(* IEC 61131-3 sources: plcassist-cli/packages/volt-lsp-iec/test-corpus/pro2193/Device/Plc Logic/Application/09 Misc/Library Manager/L_TT1P_TechnologyModules (part 3) *)

(* ---- L_MB1P_MOVEPICKANDPLACEBASE.fb ---- *)
FUNCTION_BLOCK L_MB1P_MOVEPICKANDPLACEBASE EXTENDS L_MC4P_Template_AG_KIN
VAR_INPUT
	DWCYCLESTAMP : DWORD;
	XEXECUTE : BOOL;
	XABORT : BOOL;
	WMOVEMODE : WORD;
	XFULLPATHBLENDING : BOOL;
	XNOTCOORDINATEDSTOPALL : BOOL;
	ETARGETCOORDSYSTEM : L_MC4P_CoordSystem;
	ESTARTCOORDSYSTEM : L_MC4P_CoordSystem;
	LRSTARTBLENDINGRADIUS : LREAL;
	EBUFFERMODE : MC_BUFFER_MODE := MC_BUFFER_MODE.mcBlendingLow;
	LRPATHJERK : LREAL := 1E+24;
	LRGRIPPERTIME : LREAL;
	XPULSEGRIPPERINTERRUPT : BOOL;
	XCALCPROFILEMOVEPATH : BOOL;
	WCONVEYOREXTRAPOLMODE : WORD;
	LRCONVEYOREXTRAPOLOFFSET : LREAL;
	LRCONVEYOREXTRAPOLVEL : LREAL;
	LRCONVEYOREXTRAPOLTIME : LREAL;
	XGETOVERRIDEFADINGTIME : BOOL;
END_VAR
VAR_OUTPUT
	XERROR : BOOL;
	XWARNING : BOOL;
	EERRORID : L_IE1P_Error;
	XBUSY : BOOL;
	XDONE : BOOL;
	XPROFILEINPREPARATION : BOOL;
	XCOMMANDABORTED : BOOL;
	XACTIVE : BOOL;
	XPATHHOLD : BOOL;
	XPATHHOLDONGRIPPERPOINT : BOOL;
	ESETSEGMENTTYPEOUT : L_MC4P_SegmentType;
	ALRTARGETPOSWCSOUT : ARRAY [1..6] OF LREAL;
	ALRTARGETPOSAUXOUT : ARRAY [1..6] OF LREAL;
	XPULSEGRIPPER : BOOL;
	WPATHMODEOUT : WORD;
	ITARGETPOINT : SINT;
	INUMOFSEGMENTSINPROFILE : SINT;
	XSETPATHPREPARATIONTIMEVALID : BOOL;
	LRSETPATHPREPARATIONTIMEOUT : LREAL;
	LRSETPROFILEIPOTIMEOUT : LREAL;
	XPRECALCPROFILERESTTIMEVALID : BOOL;
	LRPRECALCPROFILERESTTIME : LREAL;
	LRPRECALCPROFILEORIRESTTIME : LREAL;
	XUPDATEPROFILESYNCRESTTIME : BOOL;
	XPRECALCPROFILESYNCRESTTIME : BOOL;
	LRPRECALCPROFILESYNCRESTTIME : LREAL;
	XPRECALCPROFILESYNCOUTTIME : BOOL;
	LRPRECALCPROFILESYNCOUTTIME : LREAL;
	LRPRECALCPROFILETIME : LREAL;
	LRINTERRUPTPATHACC : LREAL;
	XIPOTIMEMOVEFROMTARGETVALID : BOOL;
	WIPOTIMEMOVEFROMTARGETCVNO : WORD;
	LRIPOTIMEMOVEFROMTARGET : LREAL;
	LRCONVEYOREXTRAPOLOFFSETOUT : LREAL;
	XPARVALID : BOOL := FALSE;
	LROVERRIDEFADINGTIME : LREAL;
	LRMAXVEL : LREAL := 10;
	LRMAXACC : LREAL := 100;
	LRMAXDEC : LREAL := 100;
	LRMAXJERK : LREAL := 100;
	XRESERVEFUNID : BOOL;
	XWAITDISABLEMOVECONTPATH : BOOL;
END_VAR
VAR_IN_OUT
	MC_MOVELINABSCONTINUEPROFILE : L_MC4P_MoveLinearAbsolute_Internal;
END_VAR
VAR
	WMOVEMODE_INT : WORD;
	XSINGLESTEP_INT : BOOL;
	XPULSEGRIPPERINTERRUPT_INT : BOOL;
	LRSTARTBLENDINGRADIUS_INT : LREAL;
	ICONTPGRIPPERINTERRUPT_INT : INT;
	XINTERRUPTONGRIPPERPOINTATMODE_INT : BOOL;
	LRPRECALCPROFILERESTTIME_INT : LREAL;
	LRSETPROFILEIPOTIME_INT : LREAL;
	LRACTTIMEOR : LREAL;
	LRSYNCRONISEDTIME : LREAL;
	LRACTSYNCRONISEDTIME : LREAL;
	XACTSYNCRONISEDTIMEOLDVALID : BOOL;
	LRACTSYNCRONISEDTIME_OLD : LREAL;
	XRESETSUPERPOSONCV_INT : BOOL;
	LRSYNCINZDISTFACTOR_INT : LREAL := 0.5;
	LRSYNCINDISTFACTOR_INT : LREAL := 1;
	LRSYNCOUTDISTFACTOR_INT : LREAL := 1;
	LRWAITTIMESTATICTARGETPOS_INT : LREAL;
	XINTERRUPTATSTATICTARGETPOS_INT : BOOL;
	XINTERRUPTATTARGETONCV_INT : BOOL;
	XABORTACTIVE : BOOL;
	WMODE_OLD : WORD;
	WMODE_INT : WORD;
	LRADDPROFILERESTTIME_INT : LREAL;
	XADDPROFILERESTTIMEVALID : BOOL;
	XACKNTARGETWORKPIECE_INT : BOOL;
	LRAUX1STARTPOS_INT : LREAL;
	XAUX1STARTPOSVALID_INT : BOOL;
	LRASTARTPOS_INT : LREAL;
	XASTARTPOSVALID_INT : BOOL;
	LRBSTARTPOS_INT : LREAL;
	XBSTARTPOSVALID_INT : BOOL;
	LRCSTARTPOS_INT : LREAL;
	XCSTARTPOSVALID_INT : BOOL;
	ETRACKPICKANDPLACETARGET_INT_OLD : L_TT1P_TrackPickAndPlaceTarget;
	ETRACKPICKANDPLACETARGET_INT : L_TT1P_TrackPickAndPlaceTarget;
	EBUFFERMODEINTERNAL_INT : MC_BUFFER_MODE := MC_BUFFER_MODE.mcBlendingLow;
	LWTCHECKSUM_INT : LWORD;
	LRTMPSTARTCOORDSYS : LREAL;
	LRPROFILERESTTIME : LREAL;
	XPRECALCGRIPPERRESTTIMEVALID : BOOL;
	LRPRECALCGRIPPERRESTTIME : LREAL;
	ETRACKPPMOVESTATUS_INT : L_TT1P_TrackPickAndPlaceTargetStatus;
	XPATHHOLD_INT : BOOL;
	XPAHTHOLDDONE_INT : BOOL;
	XPAHTHOLDDONE_LOCK : BOOL;
	REQUESTSINFO : DWORD;
	REQUESTSINFO_OLD : DWORD;
	DWRTRIG : DWORD;
	DWFTRIG : DWORD;
	LRTEMP : LREAL;
	LRTEMP2 : LREAL;
	IDX1 : SINT;
	IDX2 : SINT;
	UIDX : USINT;
	WDX : WORD;
	LRTIME_TMP : LREAL;
	LRALLPOFILETIME : LREAL;
	LRRESTTIMEENDSEGMENT_INT : LREAL;
	IDX_START : SINT;
	IDX_END : SINT;
	XINTERRUPTEDATNEXTBUFFEREDPOS_TMP : BOOL;
	WSTATE : WORD;
	WSTATE_OLD : WORD;
	XSTATEENTRY : BOOL;
	XIPOTIMEMOVEFROMTARGETVALID_OLD : BOOL;
	LRTASKCYCLE : LREAL;
	LRTASKCYCLEOR : LREAL;
	LRTASKCYCLE_INV : LREAL;
	XSTARTPATHLISTISEMPTY : BOOL;
	XCALCPATHPREPARATIONTIME : BOOL;
	XRETURNINIT : BOOL;
	LRTIMECORRFACTORATOR_INT : LREAL;
	LRPRECALCGRIPPERRESTTIMECORROR : LREAL;
	XPRECALCPROFILESYNCOUTTIME_INT : BOOL;
	INUMOFMOVEREL : SINT;
	INUMOFMOVEABS : SINT;
	INUMOFMOVEELLIPTICAL : SINT;
	XEXECUTEAFTERHALT : BOOL;
	INUMOFSEGMENTSEXECUTED : SINT;
	INUMOFMOVERELEXECUTED : SINT;
	INUMOFMOVEABSEXECUTED : SINT;
	INUMOFMOVEELLIPTICALEXECUTED : SINT;
	INUMOFMOVESPLINEEXECUTED : SINT;
	ITARGETPOINTMOVEABS : SINT;
	XNOMOVEFBEXECUTED : BOOL;
	INUMOFMOVEFBSCHECKEDORFEEDINGTIME : SINT;
	LRZSYNCDIST : LREAL;
	EPATHMODE_INT : L_TT1P_PickAndPlacePathMode;
	XGRIPPERCTRLACTIVE_INT : BOOL;
	ISETMOVEFBNOACTIVE : SINT;
	ISETNUMOFMOVEFBSADDTIME : SINT;
	IACKNNUMOFSEGMENTSINPROFILE : SINT;
	IACKNNUMOFMOVEREL : SINT;
	IACKNNUMOFMOVEABS : SINT;
	IACKNNUMOFMOVEELLIPTICAL : SINT;
	INUMOFENABLEDSEGMENTS : SINT;
	XPROFILEINPREPARATION_INT : BOOL;
	XMOVEPROFILEBUSY : BOOL;
	XMOVEPROFILEACTIVE : BOOL;
	XMOVEPROFILEACTIVE_OLD : BOOL;
	XMOVEPROFILEDONE : BOOL;
	XMOVEPROFILENOPULSEGRIPPERDONE : BOOL;
	XMOVEPROFILECOMMANDABORTED : BOOL;
	XMOVEPROFILECOMMANDABORTED_OLD : BOOL;
	XMOVEPROFILEENABLED : BOOL;
	XMOVEPROFILEHOLD : BOOL;
	XHOLDONHALT : BOOL;
	XHOLDONGRIPPERPOINT : BOOL;
	XHOLDONGRIPPERPOINT_OLD : BOOL;
	XMOVEPROFILEERROR : BOOL;
	EMOVEPROFILEERRORID : L_IE1P_Error;
	XMOVEPROFILESTATEINITIAL : BOOL := TRUE;
	ITARGETPOINTOFFSET : INT;
	INUMOFVALIDPROFILETIME : USINT;
	AXPROFILETIMEVALID : ARRAY [1..11] OF BOOL;
	ALRPROFILETIME : ARRAY [1..11] OF LREAL;
	WTARGETMODE_INT : WORD;
	XPRECALCPROFILERESTTIMEVALID_INT : BOOL;
	XPRECALCPROFILERESTTIMEVALID_OLD : BOOL;
	XCONTINUE1STMOVEABSACTIVE : BOOL;
	XCONTINUEPROFILEVIA1STMOVEABS : BOOL;
	XERROR_INVALIDCOORDSYSTEM : BOOL;
	XERRORINVALIDPROFILE : BOOL;
	XERROR_INTERNAL : BOOL;
	IINVALIDEMOVESTATECOUNTER : INT := 0;
	XSETZPOSVALID : BOOL;
	LRSETZPOSITION : LREAL;
	LRSETZPOSITION_OLD : LREAL;
	LRSETZDIST_INT : LREAL;
	LRPATHDIST_INT : LREAL;
	EBUFFERMODEINTERNAL : MC_BUFFER_MODE;
	ETRACKPICKANDPLACETARGET : L_TT1P_TrackPickAndPlaceTarget;
	ETRACKPICKANDPLACETARGET_OLD : L_TT1P_TrackPickAndPlaceTarget;
	ETRACKPPMOVESTATUS : L_TT1P_TrackPickAndPlaceTargetStatus;
	INUMOFACTIVEPATHSEGMENT : INT;
	LRADDPROFILERESTTIME : LREAL;
	LRAUX1STARTPOS : LREAL;
	LRPRECALCINGRIPPERPOSRESTTIME : LREAL;
	LRSYNCINDISTFACTOR : LREAL;
	LRSYNCINZDISTFACTOR : LREAL;
	LRSYNCOUTDISTFACTOR : LREAL;
	LRWAITTIMESTATICTARGETPOS : LREAL;
	LWTCHECKSUM : LWORD;
	WMODE : WORD;
	WMODEOLD : WORD;
	WSTATELINE : WORD;
	XACKNTARGETWORKPIECE : BOOL;
	XGRIPPERCTRLACTIVE : BOOL;
	XGRIPPERSEGMENTTIMEIPOACTIVE : BOOL;
	XINGRIPPERPOS : BOOL;
	XINTERRUPTATSTATICTARGET : BOOL;
	XINTERRUPTATTARGETONCV : BOOL;
	XLASTSEGMENTTIMEIPOACTIVE : BOOL;
	XPATHHOLDONENDHALT : BOOL;
	XPRECALCINGRIPPERPOSRESTTIMEVALID : BOOL;
	XRESETSUPERPOSONCV : BOOL;
	XRTRIGIPOTIMEMOVEFROMTARGETVALID : BOOL;
END_VAR
END_FUNCTION_BLOCK

METHOD ABORT
END_METHOD

METHOD CALL_ABORTINPUT
END_METHOD

METHOD CALL_ALLOCPOINTADR
END_METHOD

METHOD CALL_CALCTIME
END_METHOD

METHOD CALL_CHECKSTATEENTRY
END_METHOD

METHOD CALL_DISABLEMOVECONTPATH
VAR_IN_OUT
	AXESGROUP : AXES_GROUP_KIN;
END_VAR
END_METHOD

METHOD CALL_ERRORHANDLER
END_METHOD

METHOD CALL_FBMETHODS
END_METHOD

METHOD CALL_FBMETHODS_MOVEFBS
END_METHOD

METHOD CALL_GRIPPERCONTROL
END_METHOD

METHOD CALL_MC_MOVELINABS
VAR_IN_OUT
	AXESGROUP : AXES_GROUP_KIN;
END_VAR
END_METHOD

METHOD CALL_MC_MOVELINABS_1STCONTINUEPROFILE
VAR_IN_OUT
	AXESGROUP : AXES_GROUP_KIN;
END_VAR
END_METHOD

METHOD CALL_OUTPUT
END_METHOD

METHOD CALL_OUTPUTDISABLED
END_METHOD

METHOD CALL_PROFILE_STATUS
END_METHOD

METHOD CALL_PROFILE_STATUS_1STCONTINUEPROFILE
END_METHOD

METHOD CALL_PROFILE_STATUS_INIT
END_METHOD

METHOD CALL_PROFILE_STATUS_OUTPUT
END_METHOD

METHOD CALL_REQUESTS_EXT
END_METHOD

METHOD CALL_RESET
END_METHOD

METHOD CALL_RESETCOMMANDS
END_METHOD

METHOD CALL_RESETOUTPUT
END_METHOD

METHOD CALL_RESETTEMPMEMORY
END_METHOD

METHOD CALL_STATEMACHINE
END_METHOD

METHOD GET_LRPRECALCPROFILERESTTIMEFASTSYNCOUT : LREAL
END_METHOD

METHOD GET_LRRESTTIMEBEVOREMOVETOPARKPOS : LREAL
END_METHOD

METHOD GET_LRPROFILETIMEZTARGETDIST : BOOL
VAR_IN_OUT
	XPROFILETIMEZTARGETDISTVALID : BOOL;
	LRPROFILETIMEZTARGETDIST : LREAL;
END_VAR
END_METHOD

METHOD SET_EXTERNALGRIPPERTRIGGER
END_METHOD

METHOD CALL_EMPTY
END_METHOD

METHOD CALL_CONTINUEPROFILE
END_METHOD

METHOD CALL_CONTINUEPROFILE1STBLENDING
END_METHOD

METHOD CALL_CONTINUEPROFILE_MOVEABSCONTINUEPROFILE
END_METHOD

METHOD CALL_DATAFROMIPOLISTELEMENT
END_METHOD

METHOD CALL_DATAFROMIPOLISTELEMENTATSTOP
END_METHOD

METHOD CALL_DISABLEMOVEFBS
END_METHOD

METHOD CALL_EXECUTEPROFILE
END_METHOD

METHOD CALL_LOCKPAR
END_METHOD

METHOD CALL_READSTARTPOSITION
END_METHOD

METHOD CALL_SETPROFILE
END_METHOD

METHOD FUN_GETOVERRIDEFADINGTIME
VAR_INPUT
	INUMOFMOVEFBS : SINT;
END_VAR
END_METHOD

METHOD GET_PROFILETIME_MOVELINABSCONTINUEPROFILE : LREAL
END_METHOD

METHOD RESET_PRECALCPROFILETIME
END_METHOD

METHOD SET_TONEXTSEGMENTAFTERPATHHOLD
END_METHOD

METHOD CALL_INIT
END_METHOD

METHOD CALL_S000_CYCLIC
END_METHOD

(* ---- L_MB1P_MOVEPICKANDPLACEBASEEXTENDED.fb ---- *)
FUNCTION_BLOCK L_MB1P_MOVEPICKANDPLACEBASEEXTENDED EXTENDS L_MB1P_MovePickAndPlaceBase
VAR_INPUT
	ALRTARGETPOS : ARRAY [1..12] OF LREAL;
	LRZSTARTDIST : LREAL;
	LRZTARGETDIST : LREAL;
	LRVELFACTORATTARGET : LREAL := 1;
	LRACCDECFACTORATTARGET : LREAL := 1;
	XZSTARTDISTTOPARKPOS : BOOL;
	LRZSTARTDISTTOPARKPOS : LREAL;
	XZTARGETDISTFROMPARKPOS : BOOL;
	LRZTARGETDISTFROMPARKPOS : LREAL;
	LRBLENDINGRADIUS : LREAL;
	LRPATHVEL : LREAL := 10;
	LRPATHACC : LREAL := 100;
	LRPATHDEC : LREAL := 100;
	EORIENTATIONMODE : L_MC4P_Orientation_Mode := L_MC4P_Orientation_Mode.ShortestSpacialWay;
	EADIRECTION : MC_DIRECTION := MC_DIRECTION.mcShortestWay;
	EBDIRECTION : MC_DIRECTION := MC_DIRECTION.mcShortestWay;
	ECDIRECTION : MC_DIRECTION := MC_DIRECTION.mcShortestWay;
END_VAR
VAR_IN_OUT
	MC_MOVELINREL : L_MC4P_MoveLinearRelative_Internal;
	AMC_MOVELINABS : ARRAY [1..2] OF L_MC4P_MoveLinearAbsolute_Internal;
END_VAR
VAR
	LRZSTARTDIST_INT : LREAL;
	LRZTARGETDIST_INT : LREAL;
	LRZDISTELLIPTICAL_INT : LREAL;
	LRZSTARTPOSWCS_INT : LREAL;
	LRZTARGETPOSWCS_INT : LREAL;
	LRZSTARTPOSINTARGET : LREAL;
	LRZTARGETPOSINTARGET : LREAL;
	LRPRECALCPROFILETIMEINTARGETCOORDSYSTEM : LREAL;
	LRPRECALCPROFILETIMEZTARGETDIST : LREAL;
	XCALCPRECALCPROFILETIMEZTARGETDIST : BOOL := FALSE;
	WPROFILEMASK_LOCK : WORD;
	WPROFILEMODE_LOCK : WORD;
	LRZDIST_INT : LREAL;
	XLASTSEGMENTTIMEIPOACTIVE : BOOL;
END_VAR
END_FUNCTION_BLOCK

METHOD CALL_CALCTIME
END_METHOD

METHOD CALL_DISABLEMOVECONTPATH
VAR_IN_OUT
	AXESGROUP : AXES_GROUP_KIN;
END_VAR
END_METHOD

METHOD CALL_FBMETHODS_MOVEFBS
END_METHOD

METHOD CALL_MC_MOVELINABS
VAR_IN_OUT
	AXESGROUP : AXES_GROUP_KIN;
END_VAR
END_METHOD

METHOD CALL_MC_MOVELINREL
VAR_IN_OUT
	AXESGROUP : AXES_GROUP_KIN;
END_VAR
END_METHOD

METHOD CALL_OUTPUTDISABLED
END_METHOD

METHOD CALL_PROFILE_STATUS
END_METHOD

METHOD CALL_PROFILE_STATUS_MOVEABS
END_METHOD

METHOD CALL_PROFILE_STATUS_MOVEREL
END_METHOD

METHOD CALL_PROFILE_STATUS_OUTPUT
END_METHOD

METHOD CALL_RESETCOMMANDS
END_METHOD

METHOD CALL_CONTINUEPROFILE
END_METHOD

METHOD CALL_CONTINUEPROFILE_MOVEABS
END_METHOD

METHOD CALL_CONTINUEPROFILE_MOVEREL
END_METHOD

METHOD CALL_DATAFROMIPOLISTELEMENTATSTOP
END_METHOD

METHOD CALL_DISABLEMOVEFBS
END_METHOD

METHOD CALL_EXECUTEPROFILE
END_METHOD

METHOD CALL_LOCKPAR
END_METHOD

METHOD CALL_LOCKPAR_ZDIST
END_METHOD

METHOD CALL_LOCKPAR_ZSTARTDISTTOPARKPOS
END_METHOD

METHOD CALL_LOCKPAR_ZTARGETDISTFROMPARKPOS
END_METHOD

METHOD CALL_SETPROFILE
END_METHOD

METHOD CALL_SETPROFILE_TOFIRSTPOINT
END_METHOD

METHOD GET_PROFILETIME_MOVELINREL : LREAL
END_METHOD

METHOD GET_PROFILETIME_AMOVEABS : LREAL
VAR_IN_OUT
	IFBNO : SINT;
END_VAR
END_METHOD

METHOD SET_TONEXTSEGMENTAFTERPATHHOLD
END_METHOD

(* ---- L_MB1P_MOVEPICKANDPLACEELLIPTICAL.fb ---- *)
FUNCTION_BLOCK L_MB1P_MOVEPICKANDPLACEELLIPTICAL EXTENDS L_MB1P_MovePickAndPlaceBaseExtended
VAR_INPUT
	EPATHMODE : L_TT1P_PickAndPlacePathMode;
	LRZDISTELLIPTICAL : LREAL;
	XZSTARTPOSMCS : LREAL;
	LRZSTARTPOSWCS : LREAL;
	LRZTARGETPOSWCS : LREAL;
	ALRDIRECTIONTOPARKPOS : ARRAY [1..3] OF LREAL := [0, 0, 1];
	ALRDIRECTIONFROMPARKPOS : ARRAY [1..3] OF LREAL := [0, 0, 1];
END_VAR
VAR_IN_OUT
	FB_MOVEELLIPTICAL : L_MC4P_MoveEllipticalAbsolutePnP_Internal;
END_VAR
VAR
	XTEST : BOOL;
	XUSEORICAM_INT : BOOL;
	LRAUX1CAMTARGETPOS : LREAL;
	LRCCAMTARGETPOS : LREAL;
	XLASTSEGMENTTIMEIPOACTIVE : BOOL;
	XUSEORICAM : BOOL;
END_VAR
END_FUNCTION_BLOCK

METHOD CALL_DISABLEMOVECONTPATH
VAR_IN_OUT
	AXESGROUP : AXES_GROUP_KIN;
END_VAR
END_METHOD

METHOD CALL_FBMETHODS_MOVEFBS
END_METHOD

METHOD CALL_FB_MOVEELLIPTICAL
VAR_IN_OUT
	AXESGROUP : AXES_GROUP_KIN;
END_VAR
END_METHOD

METHOD CALL_OUTPUTDISABLED
END_METHOD

METHOD CALL_PROFILE_STATUS
END_METHOD

METHOD CALL_PROFILE_STATUS_MOVEELLIPTICAL
END_METHOD

METHOD CALL_RESETCOMMANDS
END_METHOD

METHOD GET_LRPROFILETIMEZTARGETDIST : BOOL
VAR_IN_OUT
	XPROFILETIMEZTARGETDISTVALID : BOOL;
	LRPROFILETIMEZTARGETDIST : LREAL;
END_VAR
END_METHOD

METHOD CALL_CONTINUEPROFILE
END_METHOD

METHOD CALL_CONTINUEPROFILE_MOVEELLIPTICAL
END_METHOD

METHOD CALL_DATAFROMIPOLISTELEMENTATSTOP
END_METHOD

METHOD CALL_DISABLEMOVEFBS
END_METHOD

METHOD CALL_EXECUTEPROFILE
END_METHOD

METHOD CALL_LOCKPAR
END_METHOD

METHOD CALL_LOCKPAR_ZDIST
END_METHOD

METHOD CALL_LOCKPAR_ZSTARTDISTTOPARKPOS
END_METHOD

METHOD CALL_LOCKPAR_ZTARGETDISTFROMPARKPOS
END_METHOD

METHOD CALL_SETPROFILE
END_METHOD

METHOD CALL_SETPROFILE_TOFIRSTPOINTEXTENDEDELLIPTICAL
END_METHOD

METHOD GET_PATHLENGTH_MOVEELLIPTICAL : LREAL
END_METHOD

METHOD GET_PROFILETIME_MOVEELLIPTICAL : LREAL
END_METHOD

(* ---- L_MB1P_MOVEPICKANDPLACESTATE.fb ---- *)
FUNCTION_BLOCK L_MB1P_MOVEPICKANDPLACESTATE EXTENDS L_MB1P_MovePickAndPlaceBase
VAR_INPUT
	XINTERRUPTONGRIPPERPOINT : BOOL;
	XSHIFTEXECUTENEXTPROFILE : BOOL;
	LRPATHPREPARATIONTIME : LREAL;
	XSTARTPOINTINHALT : BOOL;
	XHOLDMOVEPATH : BOOL;
	IPOINTNOSYNCIN : SINT;
	IPOINTNOPULSEGRIPPER : SINT;
	XACKPATHHALT : BOOL;
	XEXECUTEPROFILEAFTERGRIPPER : BOOL;
END_VAR
VAR_OUTPUT
	XPATHINTERRUPTOUT : BOOL;
	ETARGETCOORDSYSTEMOUT : L_MC4P_CoordSystem;
	ALRTARGETPOS : ARRAY [1..12] OF LREAL;
	ALRINTERMEDIANTEPOINT : ARRAY [1..12] OF LREAL;
	LRENDBLENDINGRADIUS : LREAL;
	XENDHALT : BOOL;
	XEXECUTEDPROFILEAFTERGRIPPER : BOOL;
END_VAR
VAR_IN_OUT
	ASCPROFILEPAR : ARRAY [1..10] OF L_TT1P_scProfilePar;
	AMC_MOVELINABS : ARRAY [1..10] OF L_MC4P_MoveLinearAbsolute_Internal;
END_VAR
VAR
	LRPATHPREPARATIONTIME_INT : LREAL;
	XSHIFTEXECUTENEXTPROFILE_INT : BOOL;
	XWAITOFNEXTPROFILE_INT : BOOL;
	WWAITOFNEXTPROFILECNTR : WORD;
	XNEXTPROFILEWAITFOREXECUTE_INT : BOOL;
	XEXECUTEPROFILEAFTERGRIPPER_LOCK : BOOL;
	XINTERRUPTONGRIPPERPOINT_INT : BOOL;
	XINTERRUPTONGRIPPERPOINT_OLD : BOOL;
	XINGRIPPERPOS_INT : BOOL;
	XINSYNCPOS_INT : BOOL;
	LRENDPATHVEL_INT : LREAL;
	LRENDPATHACC_INT : LREAL;
	LRENDPATHDEC_INT : LREAL;
	INUMOFMOVEABSEXECUTEDAFTERHALT : SINT;
	IRETURNINITCNTR : INT;
	XREADSTARTPOSACTIVE : BOOL;
	XIPOTIMEMOVEFROMTARGETACTIVE_INT : BOOL;
	ICNTRACKPATHHALT_INT : INT;
	ICNTRACKPATHHALTREST_INT : INT;
	ICNTRACKPATHHALTFORGRIPPER_INT : INT;
	ICNTRACKPATHHALT_LOCK : INT;
	INUMOFHALTINPROFILE_INT : INT;
	IPOINTNOSYNCOUT_INT : SINT;
	IPOINTNOSYNCIN_INT : SINT;
	IPOINTNOPULSEGRIPPER_INT : SINT;
	ALRSTARTPOS_INT : ARRAY [1..6] OF LREAL;
	ECOORDSYSTEMP1START : L_MC4P_CoordSystem;
	ECOORDSYSTEMP2ACT : L_MC4P_CoordSystem;
	ECOORDSYSTEMP3NEXT : L_MC4P_CoordSystem;
	ALRP1START : ARRAY [1..3] OF LREAL;
	ALRP2ACT : ARRAY [1..3] OF LREAL;
	ALRP3NEXT : ARRAY [1..3] OF LREAL;
	XPOINTSONASTRAIGHTLINE : BOOL;
	XNOFUNKTION : BOOL;
	XSTARTPOSVALID_INT : BOOL;
	XPROFILEEXECUTED_INT : BOOL;
	XEXECUTENEXTMOVEPP_INT : BOOL;
	XACKENDHALT_INT : BOOL;
	AXHALT : ARRAY [0..10] OF BOOL;
	AITARGETPOINTOFFSETATMOVEABS : ARRAY [0..10] OF INT;
	AXMOVELINABSACTIVE : ARRAY [0..10] OF BOOL;
	XVALIDSYNCRESTTIME_OLD : BOOL;
	XVALIDSYNCRESTTIME_INT : BOOL;
	XVALIDSYNCOUTRESTTIME_OLD : BOOL;
	XVALIDSYNCOUTRESTTIME_INT : BOOL;
	LRRESTTIMESYNC_INT : LREAL;
	LRRESTTIMESYNCOUT_INT : LREAL;
	XVALIDPULSEGRIPPERRESTTIME_OLD : BOOL;
	XVALIDPULSEGRIPPERRESTTIME_INT : BOOL;
	LRPULSEGRIPPERRESTTIME_INT : LREAL;
	LRBLENDINGRADIUS_TMP : LREAL;
	XCALCDIST_TMP : BOOL;
	XCALCINTERMEDIANTEPOINT : BOOL;
	AXCALCPATHLEGTHBETWEENPOINTS : ARRAY [0..10] OF BOOL;
	ALRPATHLENGTHBETWEENPOINTS : ARRAY [0..10] OF LREAL;
	ALRAUX1POINTS : ARRAY [0..10] OF LREAL;
	ALRAPOINTS : ARRAY [0..10] OF LREAL;
	ALRBPOINTS : ARRAY [0..10] OF LREAL;
	ALRCPOINTS : ARRAY [0..10] OF LREAL;
	IFORCNT : SINT;
	XCALC999AUX1TARGETPOS : BOOL;
	XCALC999ATARGETPOS : BOOL;
	XCALC999BTARGETPOS : BOOL;
	XCALC999CTARGETPOS : BOOL;
	IFIRSTPOINTATPROFILEPAR : SINT;
	ILISTELEMENTATSTOPCNTR_INT : SINT;
	XNEXTPROFILEPOINTATBLENDING_INT : BOOL;
	MC_GROUPREADACTUALPOSITION1 : MC_GroupReadActualPosition;
	ALRPROFILESTARTPOS : ARRAY [1..6] OF LREAL;
	ILISTELEMENTATSTOPCNTR : SINT;
	LRENDPATHACC : LREAL;
	LRENDPATHDEC : LREAL;
	LRENDPATHVEL : LREAL;
	WSTATELINE : WORD;
	XEXECUTENEXTMOVEPP : BOOL;
	XGRIPPERSEGMENTTIMEIPOACTIVE : BOOL;
	XINGRIPPERPOS : BOOL;
	XLASTSEGMENTTIMEIPOACTIVE : BOOL;
	XMOVEFROMTARGETACTIVE : BOOL;
	XNEXTPROFILEPOINTATBLENDING : BOOL;
	XNEXTPROFILEWAITFOREXECUTE : BOOL;
	XPATHHOLDONENDHALT : BOOL;
END_VAR
END_FUNCTION_BLOCK

METHOD CALL_ABORTINPUT
END_METHOD

METHOD CALL_CALCTIME
END_METHOD

METHOD CALL_DISABLEMOVECONTPATH
VAR_IN_OUT
	AXESGROUP : AXES_GROUP_KIN;
END_VAR
END_METHOD

METHOD CALL_ERRORHANDLER
END_METHOD

METHOD CALL_FBMETHODS
END_METHOD

METHOD CALL_FBMETHODS_MOVEFBS
END_METHOD

METHOD CALL_MC_GROUPREADACTUALPOSITION
END_METHOD

METHOD CALL_MC_MOVELINABS
VAR_IN_OUT
	AXESGROUP : AXES_GROUP_KIN;
END_VAR
END_METHOD

METHOD CALL_OUTPUT
END_METHOD

METHOD CALL_OUTPUTDISABLED
END_METHOD

METHOD CALL_PROFILE_STATUS
END_METHOD

METHOD CALL_PROFILE_STATUS_MOVEABS
END_METHOD

METHOD CALL_PROFILE_STATUS_INIT
END_METHOD

METHOD CALL_PROFILE_STATUS_OUTPUT
END_METHOD

METHOD CALL_REQUESTS_EXT
END_METHOD

METHOD CALL_RESETCOMMANDS
END_METHOD

METHOD CALL_RESETOUTPUT
END_METHOD

METHOD GET_LRPRECALCPROFILERESTTIMEFASTSYNCOUT : LREAL
END_METHOD

METHOD GET_LRRESTTIMEBEVOREMOVETOPARKPOS : LREAL
END_METHOD

METHOD GET_IACKPATHHALTCNTRREST
VAR_IN_OUT
	ICOUNTER : INT;
END_VAR
END_METHOD

METHOD CALL_CALC999TARGETPOS
VAR_INPUT
	IPOINTNO : SINT;
END_VAR
VAR_IN_OUT
	ALRPOINTS : ARRAY [0..10] OF LREAL;
	ALRLEGTHBETWEENPOINTS : ARRAY [0..10] OF LREAL;
END_VAR
END_METHOD

METHOD CALL_CHECKORIDIRECTION_SWITCHTOSHORTESTWAY
VAR_INPUT
	LRCYCLELENGTH : LREAL;
	LRPOSSTART : LREAL;
	LRPOSEND : LREAL;
	EDIRECTION : MC_DIRECTION;
END_VAR
VAR_OUTPUT
	EDIRECTIONOUT : MC_DIRECTION;
END_VAR
END_METHOD

METHOD CALL_CONTINUEPROFILE
END_METHOD

METHOD CALL_CONTINUEPROFILE_MOVEABS
END_METHOD

METHOD CALL_DATAFROMIPOLISTELEMENTATSTOP
END_METHOD

METHOD CALL_DISABLEMOVEFBS
END_METHOD

METHOD CALL_EXECUTEPROFILE
END_METHOD

METHOD CALL_LOCKPAR
END_METHOD

METHOD CALL_READSTARTPOSITION
END_METHOD

METHOD CALL_SETPROFILE
END_METHOD

METHOD FUN_POINTSONASTRAIGHTLINE : BOOL
VAR_OUTPUT
	XNOFUNKTION : BOOL;
END_VAR
VAR_IN_OUT
	AXESGROUP : AXES_GROUP_KIN;
	ALRP1 : ARRAY [1..3] OF LREAL;
	ECOORDSYSTEMP1 : L_MC4P_CoordSystem;
	ALRP2 : ARRAY [1..3] OF LREAL;
	ECOORDSYSTEMP2 : L_MC4P_CoordSystem;
	ALRP3 : ARRAY [1..3] OF LREAL;
	ECOORDSYSTEMP3 : L_MC4P_CoordSystem;
END_VAR
END_METHOD

METHOD GET_FIRSTPROFILEPOINTPAR
VAR_IN_OUT
	SCPROFILEPAR : L_TT1P_scProfilePar;
END_VAR
END_METHOD

METHOD GET_INUMOFACTIVEHALTPOINTS : INT
END_METHOD

METHOD GET_PROFILETIME_AMOVEABS : LREAL
VAR_IN_OUT
	IFBNO : SINT;
END_VAR
END_METHOD

METHOD SET_ACKENDHALT
END_METHOD

METHOD SET_FIRSTPROFILEPOINTATBLENDING
VAR_IN_OUT
	ALRTARGETPOS : ARRAY [1..12] OF LREAL;
END_VAR
END_METHOD

METHOD SET_TONEXTSEGMENTAFTERPATHHOLD
END_METHOD

METHOD SET_ISTARTACKPATHHALTCNTR
VAR_IN_OUT
	ICOUNTER : INT;
END_VAR
END_METHOD

METHOD SET_XNEXTPROFILEWAITFOREXECUTE
END_METHOD

METHOD CALL_INIT
END_METHOD

METHOD CALL_S000_CYCLIC
END_METHOD

(* ---- L_MB1P_MULTICAMSEQUENCER.fb ---- *)
FUNCTION_BLOCK L_MB1P_MULTICAMSEQUENCER
VAR_INPUT
	XENABLE : BOOL;
	XCAMSEQUENCER : BOOL;
	EMODE : L_MB1P_CamSequenceMode;
	XCAMCHANGEINSTANT : BOOL;
	ESETCAMTABLE : L_MB1P_CamTable;
	XENDOFPROFILEIN : BOOL;
	CAMTABLE1 : MC_CAM_REF;
	CAMTABLE2 : MC_CAM_REF;
	CAMTABLE3 : MC_CAM_REF;
	CAMTABLE4 : MC_CAM_REF;
END_VAR
VAR_OUTPUT
	XDONE : BOOL;
	XBUSY : BOOL;
	XERROR : BOOL;
	EERRORID : L_IE1P_Error;
	ESETCAMTABLEOUT : L_MB1P_CamTable;
	CAMTABLEOUT : MC_CAM_REF;
END_VAR
VAR
	EFMSTATE : L_MB1P_States := L_MB1P_States.INIT;
	XINITSTATE : BOOL;
	XENABLE_OLD : BOOL;
	XLOADCAMTABLE_OLD : BOOL;
	XENDOFPROFILEIN_OLD : BOOL;
	XCAMSEQUENCER_OLD : BOOL;
	XCAMCHANGEINSTANT_OLD : BOOL;
	XCAMSEQUENCERACTIVE : BOOL;
END_VAR
END_FUNCTION_BLOCK

METHOD CALL_ERRORHANDLER
END_METHOD

METHOD CALL_FBMETHODS
END_METHOD

METHOD CALL_OUTPUT
END_METHOD

METHOD CALL_RESETCOMMANDS
END_METHOD

METHOD CALL_RESETOUTPUT
END_METHOD

METHOD CALL_STATEMACHINE
END_METHOD

METHOD CALL_SETCAMTABLEOUT
VAR_INPUT
	ESETCAMTABLE : L_MB1P_CamTable;
END_VAR
END_METHOD

METHOD CAMREFCHANGED : BOOL
VAR_IN_OUT
	CAMREFNEW : MC_CAM_REF;
	CAMREFOLD : MC_CAM_REF;
END_VAR
END_METHOD

METHOD CALL_S000_CYCLIC
END_METHOD

METHOD CALL_S001_INIT
END_METHOD

METHOD CALL_S002_READY
END_METHOD

METHOD CALL_S151_SEQUENCE_CYCLICCAM1
END_METHOD

METHOD CALL_S152_SEQUENCE_CYCLICCAM3
END_METHOD

METHOD CALL_S153_SEQUENCE_CAM1CYCLICCAM3CAM1
END_METHOD

METHOD CALL_S154_SEQUENCE_CAM1CAM2CYCLICCAM3CAM4CAM1
END_METHOD

(* ---- L_MB1P_POSPROFILER.fb ---- *)
FUNCTION_BLOCK L_MB1P_POSPROFILER
VAR_INPUT
	XEXECUTE : BOOL;
	XAUXEXECUTE : BOOL;
	XABORT : BOOL;
	XPOSMODE : BOOL;
	ROVERRIDESPEED : REAL;
	ROVERRIDEACC : REAL;
	ROVERRIDEDEC : REAL;
	ROVERRIDEJERKACC : REAL;
	ROVERRIDEJERKDEC : REAL;
	LRACTPOS : LREAL;
	LRACTSPEED : LREAL;
	LRACTACC : LREAL;
	RTASKCYCLE : REAL;
END_VAR
VAR_OUTPUT
	XBUSY : BOOL;
	XDONE : BOOL;
	XABORTED : BOOL;
	XERROR : BOOL;
	LRSETPOS : LREAL;
	LRSETSPEED : LREAL;
	LRSETACC : LREAL;
	DWSTATE : DWORD;
	DWPROFILETYPE : DWORD;
END_VAR
VAR_IN_OUT
	SCPROFILEPARAMETER : L_MB1P_ProfileParameter;
END_VAR
VAR
	SCPROFILEDATA : L_MB1P_ProfileData;
	LREVALTIME : LREAL;
	DWSTATEOFINTERPOLATOR : DWORD;
	XFLAGEXECUTE : BOOL;
	XFLAGAUXEXECUTE : BOOL;
	XFLAGABORT : BOOL;
	SCPROFILEPARAMETERINT : L_MB1P_ProfileParameter;
	ROVERRIDESPEEDOLD : REAL;
	ROVERRIDEACCOLD : REAL;
	ROVERRIDEDECOLD : REAL;
	ROVERRIDEJERKACCOLD : REAL;
	ROVERRIDEJERKDECOLD : REAL;
	XSTARTCALCPROF : BOOL;
	XVELOVEREQZERO : BOOL;
	ARG1 : LREAL;
END_VAR
END_FUNCTION_BLOCK

METHOD CALCPROFILE : BOOL
VAR_INPUT
	DWPROFILETYPE : DWORD;
	LRSTARTACC : LREAL;
	LRSTARTVEL : LREAL;
	SCPROFILEPARAMETER : L_MB1P_ProfileParameter;
	SCMINPROFILEDATA : L_MB1P_IntProfileData;
	SCMAXPROFILEDATA : L_MB1P_IntProfileData;
END_VAR
VAR_OUTPUT
	SCPROFILEDATA : L_MB1P_ProfileData;
	DWSTATE : DWORD;
END_VAR
END_METHOD

METHOD CALCPROFILEDATA : BOOL
VAR_INPUT
	LRSTARTACC : LREAL;
	LRSTARTVEL : LREAL;
	LRSTARTPOS : LREAL;
	XVELMODE : BOOL;
END_VAR
VAR_OUTPUT
	XERROR : BOOL;
	DWSTATE : DWORD;
	DWPROFILETYPE : DWORD;
END_VAR
VAR_IN_OUT
	SCPROFILEDATA : L_MB1P_ProfileData;
	SCPROFILEPARAMETER : L_MB1P_ProfileParameter;
END_VAR
END_METHOD

METHOD IDENTPROFILETYPE : DWORD
VAR_INPUT
	XVELMODE : BOOL;
	LRSTARTACC : LREAL;
	LRSTARTVEL : LREAL;
	SCPROFILEPARAMETER : L_MB1P_ProfileParameter;
END_VAR
VAR_OUTPUT
	DWPROFILETYPE : DWORD;
	SCMINPROFILEDATA : L_MB1P_IntProfileData;
	SCMAXPROFILEDATA : L_MB1P_IntProfileData;
	DWSTATE : DWORD;
END_VAR
END_METHOD

METHOD PROFILEINTERPOLATOR : BOOL
VAR_INPUT
	LREVALTIME : LREAL;
END_VAR
VAR_OUTPUT
	DWSTATE : DWORD;
	LRSETPOS : LREAL;
	LRSETVEL : LREAL;
	LRSETACC : LREAL;
END_VAR
VAR_IN_OUT
	SCPROFILEDATA : L_MB1P_ProfileData;
END_VAR
END_METHOD

METHOD RESETOUTPUT
END_METHOD

METHOD CALCSQRT : LREAL
VAR_INPUT
	ARG1 : LREAL;
END_VAR
END_METHOD

METHOD CALCMINPOSPROFILE : BOOL
VAR_INPUT
	MAXVEL : LREAL;
	MAXACC1 : LREAL;
	MAXACC2 : LREAL;
	JERKACC1 : LREAL;
	JERKACC2 : LREAL;
	RECIPRJERKACC1 : LREAL;
	RECIPRJERKACC2 : LREAL;
	V0_ACC1 : LREAL;
	V0_ACC2 : LREAL;
	A0_ACC1 : LREAL;
	A0_ACC2 : LREAL;
END_VAR
VAR_OUTPUT
	DIMINPOSPROFILETYPE : DINT;
	MINPOSPROFILEDATA : L_MB1P_IntProfileData;
	VMAXMINTRIACC1 : LREAL;
	VMAX_MINTRIACC2 : LREAL;
END_VAR
END_METHOD

METHOD CALCMINPROFILENEGACC : BOOL
VAR_INPUT
	VMAX : LREAL;
	AMAX : LREAL;
	V0 : LREAL;
	A0 : LREAL;
	JERK : LREAL;
	JERKRECIPR : LREAL;
END_VAR
VAR_OUTPUT
	DWPROFILETYPE : DWORD;
	PROFILEDATA_NEGACC : L_MB1P_IntProfileDataAcc;
END_VAR
END_METHOD

METHOD CALCMINPROFILEPOSACC : BOOL
VAR_INPUT
	VMAX : LREAL;
	AMAX : LREAL;
	V0 : LREAL;
	A0 : LREAL;
	JERK : LREAL;
	JERKRECIPR : LREAL;
END_VAR
VAR_OUTPUT
	DWPROFILETYPE : DWORD;
	PROFILEDATA_POSACC : L_MB1P_IntProfileDataAcc;
END_VAR
END_METHOD

METHOD CALCMINTRI : BOOL
VAR_INPUT
	RECIPRJERKACC1 : LREAL;
	RECIPRJERKACC2 : LREAL;
	A0_ACC1 : LREAL;
	V0_ACC1 : LREAL;
	A0_ACC2 : LREAL;
	V0_ACC2 : LREAL;
END_VAR
VAR_OUTPUT
	VMAXMINTRIACC1 : LREAL;
	VMAXMINTRIACC2 : LREAL;
	PROFILEDATA_ACC1 : L_MB1P_IntProfileDataAcc;
	PROFILEDATA_ACC2 : L_MB1P_IntProfileDataAcc;
END_VAR
END_METHOD

METHOD CHECKPROFILEDATA
VAR_INPUT
	DWMODE : DWORD;
	LRTARGETPOS : LREAL;
	LRTARGETVEL : LREAL;
	LRTARGETACC : LREAL;
	LRJERKPHASE7 : LREAL;
END_VAR
VAR_OUTPUT
	XERROR : BOOL;
END_VAR
VAR_IN_OUT
	SCPROFILEDATA : L_MB1P_ProfileData;
END_VAR
END_METHOD

METHOD IDENTMINNEGPROFILE : BOOL
VAR_INPUT
	MINPOSPROFILETYPE : DINT;
	MAXVEL : LREAL;
	MAXACC : LREAL;
	JERK : LREAL;
	RECIPRJERK : LREAL;
	V0_ACC1 : LREAL;
	V0_ACC2 : LREAL;
	A0_ACC1 : LREAL;
	A0_ACC2 : LREAL;
	TARGETPOS : LREAL;
END_VAR
VAR_OUTPUT
	DWPROFILETYPE : DWORD;
END_VAR
VAR_IN_OUT
	SCMAXPROFILEDATA : L_MB1P_IntProfileData;
	SCMINPROFILEDATA : L_MB1P_IntProfileData;
END_VAR
END_METHOD

METHOD IDENTMINPOSPROFILE : BOOL
VAR_INPUT
	MAXVEL : LREAL;
	MAXACC1 : LREAL;
	MAXACC2 : LREAL;
	JERKACC1 : LREAL;
	JERKACC2 : LREAL;
	V0_ACC1 : LREAL;
	V0_ACC2 : LREAL;
	A0_ACC1 : LREAL;
	A0_ACC2 : LREAL;
	TARGETPOS : LREAL;
END_VAR
VAR_OUTPUT
	DWPROFILETYPE : DWORD;
	SCMAXPROFILEDATA : L_MB1P_IntProfileData;
	SCMINPROFILEDATA : L_MB1P_IntProfileData;
END_VAR
END_METHOD

METHOD IDENTSIMPLETRAPNEG : BOOL
VAR_INPUT
	MAXACC2 : LREAL;
	V0_ACC1 : LREAL;
	V0_ACC2 : LREAL;
	A0_ACC1 : LREAL;
	A0_ACC2 : LREAL;
	JERKACC1 : LREAL;
	JERKACC2 : LREAL;
	RECIPRJERKACC2 : LREAL;
	TARGETPOS : LREAL;
END_VAR
VAR_OUTPUT
	DWPROFILETYPE : DWORD;
END_VAR
VAR_IN_OUT
	SCMINPROFILEDATA : L_MB1P_IntProfileData;
	SCMAXPROFILEDATA : L_MB1P_IntProfileData;
END_VAR
END_METHOD

METHOD IDENTSIMPLETRAPPOSTRINEG : BOOL
VAR_INPUT
	MAXACC1 : LREAL;
	JERKACC1 : LREAL;
	RECIPRJERKACC1 : LREAL;
	V0_ACC1 : LREAL;
	A0_ACC1 : LREAL;
	VMAXMINTRIACC1 : LREAL;
	VMAXMINTRIACC2 : LREAL;
	JERKACC2 : LREAL;
	TARGETPOS : LREAL;
END_VAR
VAR_OUTPUT
	DWPROFILETYPE : DWORD;
END_VAR
VAR_IN_OUT
	SCMINPROFILEDATA : L_MB1P_IntProfileData;
	SCMAXPROFILEDATA : L_MB1P_IntProfileData;
END_VAR
END_METHOD

METHOD IDENTSIMPLETRINEG : BOOL
VAR_INPUT
	V0_ACC1 : LREAL;
	A0_ACC1 : LREAL;
	A0_ACC2 : LREAL;
	JERKACC1 : LREAL;
	JERKACC2 : LREAL;
	RECIPRJERKACC2 : LREAL;
	TARGETPOS : LREAL;
END_VAR
VAR_OUTPUT
	DWPROFILETYPE : DWORD;
END_VAR
VAR_IN_OUT
	SCMINPROFILEDATA : L_MB1P_IntProfileData;
	SCMAXPROFILEDATA : L_MB1P_IntProfileData;
END_VAR
END_METHOD

METHOD IDENTSIMPLETRIPOSTRAPNEG : BOOL
VAR_INPUT
	MAXACC2 : LREAL;
	JERKACC2 : LREAL;
	RECIPRJERKACC2 : LREAL;
	V0_ACC2 : LREAL;
	A0_ACC2 : LREAL;
	VMAXMINTRIACC1 : LREAL;
	JERKACC1 : LREAL;
	TARGETPOS : LREAL;
END_VAR
VAR_OUTPUT
	DWPROFILETYPE : DWORD;
END_VAR
VAR_IN_OUT
	SCMINPROFILEDATA : L_MB1P_IntProfileData;
	SCMAXPROFILEDATA : L_MB1P_IntProfileData;
END_VAR
END_METHOD

METHOD IDENTSIMPLETRIPOSTRINEG : BOOL
VAR_INPUT
	V0_ACC1 : LREAL;
	A0_ACC1 : LREAL;
	AMAX : LREAL;
	RECIPRJERKACC1 : LREAL;
	JERKACC1 : LREAL;
	JERKACC2 : LREAL;
	TARGETPOS : LREAL;
	VMAXMINTRIACC1 : LREAL;
	VMAXMINTRIACC2 : LREAL;
END_VAR
VAR_OUTPUT
	DWPROFILETYPE : DWORD;
END_VAR
VAR_IN_OUT
	SCMINPROFILEDATA : L_MB1P_IntProfileData;
	SCMAXPROFILEDATA : L_MB1P_IntProfileData;
END_VAR
END_METHOD

METHOD IDENTTRAPTRI : BOOL
VAR_INPUT
	V_MINTRAPEZACC1 : LREAL;
	MAXACC1 : LREAL;
	JERKACC1 : LREAL;
	JERKACC2 : LREAL;
	A0_ACC1 : LREAL;
	A0_ACC2 : LREAL;
	V0_ACC1 : LREAL;
	V0_ACC2 : LREAL;
	T1_ACC1 : LREAL;
	T3_ACC1 : LREAL;
	DS_1_ACC1 : LREAL;
	TARGETPOS : LREAL;
END_VAR
VAR_OUTPUT
	DWPROFILETYPE : DWORD;
END_VAR
VAR_IN_OUT
	SCMINPROFILEDATA : L_MB1P_IntProfileData;
	SCMAXPROFILEDATA : L_MB1P_IntProfileData;
END_VAR
END_METHOD

METHOD IDENTTRITRAP : BOOL
VAR_INPUT
	V_MINTRAPEZACC2 : LREAL;
	MAXACC2 : LREAL;
	JERKACC1 : LREAL;
	JERKACC2 : LREAL;
	A0_ACC1 : LREAL;
	A0_ACC2 : LREAL;
	V0_ACC1 : LREAL;
	V0_ACC2 : LREAL;
	T1_ACC2 : LREAL;
	T3_ACC2 : LREAL;
	DS_1_ACC2 : LREAL;
	TARGETPOS : LREAL;
END_VAR
VAR_OUTPUT
	DWPROFILETYPE : DWORD;
END_VAR
VAR_IN_OUT
	SCMINPROFILEDATA : L_MB1P_IntProfileData;
	SCMAXPROFILEDATA : L_MB1P_IntProfileData;
END_VAR
END_METHOD

METHOD CALCPROFILE_10A0 : BOOL
VAR_INPUT
	LRSTARTACC : LREAL;
	LRSTARTVEL : LREAL;
	LRMAXACC : LREAL;
	LRMAXDEC : LREAL;
	LRMAXVEL : LREAL;
	LRTARGETACC : LREAL;
	LRTARGETVEL : LREAL;
	LRTARGETPOS : LREAL;
	LRJERKACC : LREAL;
	LRJERKDEC : LREAL;
	LRJERKTIMEACC : LREAL;
	LRJERKTIMEDEC : LREAL;
END_VAR
VAR_OUTPUT
	DWSTATE : DWORD;
END_VAR
VAR_IN_OUT
	SCPROFILEDATA : L_MB1P_ProfileData;
	SCPROFILEPARAMETER : L_MB1P_ProfileParameter;
END_VAR
END_METHOD

METHOD CALCPROFILE_10A0_A0GTAMAX : BOOL
VAR_INPUT
	LRSTARTACC : LREAL;
	LRSTARTVEL : LREAL;
	LRMAXACC : LREAL;
	LRMAXVEL : LREAL;
	LRMAXDEC : LREAL;
	LRTARGETACC : LREAL;
	LRTARGETVEL : LREAL;
	LRTARGETPOS : LREAL;
	LRJERKTIMEACC : LREAL;
	LRJERKTIMEDEC : LREAL;
	LRJERKACC : LREAL;
	LRJERKDEC : LREAL;
END_VAR
VAR_IN_OUT
	SCPROFILEDATA : L_MB1P_ProfileData;
END_VAR
END_METHOD

METHOD CALCPROFILE_10A0_A0LTAMAX : BOOL
VAR_INPUT
	LRSTARTACC : LREAL;
	LRSTARTVEL : LREAL;
	LRMAXACC : LREAL;
	LRMAXVEL : LREAL;
	LRMAXDEC : LREAL;
	LRTARGETACC : LREAL;
	LRTARGETVEL : LREAL;
	LRTARGETPOS : LREAL;
	LRJERKTIMEACC : LREAL;
	LRJERKTIMEDEC : LREAL;
	LRJERKACC : LREAL;
	LRJERKDEC : LREAL;
END_VAR
VAR_IN_OUT
	SCPROFILEDATA : L_MB1P_ProfileData;
END_VAR
END_METHOD

METHOD CALCPROFILE_10B0 : BOOL
VAR_INPUT
	LRSTARTACC : LREAL;
	LRSTARTVEL : LREAL;
	LRMAXACC : LREAL;
	LRMAXDEC : LREAL;
	LRMAXVEL : LREAL;
	LRTARGETACC : LREAL;
	LRTARGETVEL : LREAL;
	LRTARGETPOS : LREAL;
	LRJERKACC : LREAL;
	LRJERKDEC : LREAL;
	LRJERKTIMEACC : LREAL;
	LRJERKTIMEDEC : LREAL;
END_VAR
VAR_OUTPUT
	DWSTATE : DWORD;
END_VAR
VAR_IN_OUT
	SCPROFILEDATA : L_MB1P_ProfileData;
	SCPROFILEPARAMETER : L_MB1P_ProfileParameter;
END_VAR
END_METHOD

METHOD CALCPROFILE_10B0_A0GTAMAX : BOOL
VAR_INPUT
	LRSTARTACC : LREAL;
	LRSTARTVEL : LREAL;
	LRMAXACC : LREAL;
	LRMAXVEL : LREAL;
	LRMAXDEC : LREAL;
	LRTARGETACC : LREAL;
	LRTARGETVEL : LREAL;
	LRTARGETPOS : LREAL;
	LRJERKTIMEACC : LREAL;
	LRJERKTIMEDEC : LREAL;
	LRJERKACC : LREAL;
	LRJERKDEC : LREAL;
END_VAR
VAR_IN_OUT
	SCPROFILEDATA : L_MB1P_ProfileData;
END_VAR
END_METHOD

METHOD CALCPROFILE_10B0_A0LTAMAX : BOOL
VAR_INPUT
	LRSTARTACC : LREAL;
	LRSTARTVEL : LREAL;
	LRMAXACC : LREAL;
	LRMAXVEL : LREAL;
	LRMAXDEC : LREAL;
	LRTARGETACC : LREAL;
	LRTARGETVEL : LREAL;
	LRTARGETPOS : LREAL;
	LRJERKTIMEACC : LREAL;
	LRJERKTIMEDEC : LREAL;
	LRJERKACC : LREAL;
	LRJERKDEC : LREAL;
END_VAR
VAR_IN_OUT
	SCPROFILEDATA : L_MB1P_ProfileData;
END_VAR
END_METHOD

METHOD CALCPROFILE_10C0 : BOOL
VAR_INPUT
	LRSTARTACC : LREAL;
	LRSTARTVEL : LREAL;
	LRMAXACC : LREAL;
	LRMAXDEC : LREAL;
	LRMAXVEL : LREAL;
	LRTARGETACC : LREAL;
	LRTARGETVEL : LREAL;
	LRTARGETPOS : LREAL;
	LRJERKACC : LREAL;
	LRJERKDEC : LREAL;
	LRJERKTIMEACC : LREAL;
	LRJERKTIMEDEC : LREAL;
END_VAR
VAR_OUTPUT
	DWSTATE : DWORD;
END_VAR
VAR_IN_OUT
	SCPROFILEDATA : L_MB1P_ProfileData;
	SCPROFILEPARAMETER : L_MB1P_ProfileParameter;
END_VAR
END_METHOD

METHOD CALCPROFILE_10C0_A0LTAMAXT31 : BOOL
VAR_INPUT
	LRSTARTACC : LREAL;
	LRSTARTVEL : LREAL;
	LRMAXACC : LREAL;
	LRMAXVEL : LREAL;
	LRMAXDEC : LREAL;
	LRTARGETACC : LREAL;
	LRTARGETVEL : LREAL;
	LRTARGETPOS : LREAL;
	LRJERKTIMEACC : LREAL;
	LRJERKTIMEDEC : LREAL;
	LRJERKACC : LREAL;
	LRJERKDEC : LREAL;
END_VAR
VAR_IN_OUT
	SCPROFILEDATA : L_MB1P_ProfileData;
END_VAR
END_METHOD

METHOD CALCPROFILE_10C0_A0LTAMAXT32 : BOOL
VAR_INPUT
	LRSTARTACC : LREAL;
	LRSTARTVEL : LREAL;
	LRMAXACC : LREAL;
	LRMAXVEL : LREAL;
	LRMAXDEC : LREAL;
	LRTARGETACC : LREAL;
	LRTARGETVEL : LREAL;
	LRTARGETPOS : LREAL;
	LRJERKTIMEACC : LREAL;
	LRJERKTIMEDEC : LREAL;
	LRJERKACC : LREAL;
	LRJERKDEC : LREAL;
END_VAR
VAR_IN_OUT
	SCPROFILEDATA : L_MB1P_ProfileData;
END_VAR
END_METHOD

METHOD CALCPROFILE_10D0 : BOOL
VAR_INPUT
	LRSTARTACC : LREAL;
	LRSTARTVEL : LREAL;
	LRMAXACC : LREAL;
	LRMAXDEC : LREAL;
	LRMAXVEL : LREAL;
	LRTARGETACC : LREAL;
	LRTARGETVEL : LREAL;
	LRTARGETPOS : LREAL;
	LRJERKACC : LREAL;
	LRJERKDEC : LREAL;
	LRJERKTIMEACC : LREAL;
	LRJERKTIMEDEC : LREAL;
END_VAR
VAR_OUTPUT
	DWSTATE : DWORD;
END_VAR
VAR_IN_OUT
	SCPROFILEDATA : L_MB1P_ProfileData;
	SCPROFILEPARAMETER : L_MB1P_ProfileParameter;
END_VAR
END_METHOD

METHOD CALCPROFILE_10D0_A0LTAMAXT31T51 : BOOL
VAR_INPUT
	LRSTARTACC : LREAL;
	LRSTARTVEL : LREAL;
	LRMAXACC : LREAL;
	LRMAXVEL : LREAL;
	LRMAXDEC : LREAL;
	LRTARGETACC : LREAL;
	LRTARGETVEL : LREAL;
	LRTARGETPOS : LREAL;
	LRJERKTIMEACC : LREAL;
	LRJERKTIMEDEC : LREAL;
	LRJERKACC : LREAL;
	LRJERKDEC : LREAL;
END_VAR
VAR_IN_OUT
	SCPROFILEDATA : L_MB1P_ProfileData;
END_VAR
END_METHOD

METHOD CALCPROFILE_10D0_A0LTAMAXT31T52 : BOOL
VAR_INPUT
	LRSTARTACC : LREAL;
	LRSTARTVEL : LREAL;
	LRMAXACC : LREAL;
	LRMAXVEL : LREAL;
	LRMAXDEC : LREAL;
	LRTARGETACC : LREAL;
	LRTARGETVEL : LREAL;
	LRTARGETPOS : LREAL;
	LRJERKTIMEACC : LREAL;
	LRJERKTIMEDEC : LREAL;
	LRJERKACC : LREAL;
	LRJERKDEC : LREAL;
END_VAR
VAR_IN_OUT
	SCPROFILEDATA : L_MB1P_ProfileData;
END_VAR
END_METHOD

METHOD CALCPROFILE_10D0_A0LTAMAXT32T51 : BOOL
VAR_INPUT
	LRSTARTACC : LREAL;
	LRSTARTVEL : LREAL;
	LRMAXACC : LREAL;
	LRMAXVEL : LREAL;
	LRMAXDEC : LREAL;
	LRTARGETACC : LREAL;
	LRTARGETVEL : LREAL;
	LRTARGETPOS : LREAL;
	LRJERKTIMEACC : LREAL;
	LRJERKTIMEDEC : LREAL;
	LRJERKACC : LREAL;
	LRJERKDEC : LREAL;
END_VAR
VAR_IN_OUT
	SCPROFILEDATA : L_MB1P_ProfileData;
END_VAR
END_METHOD

METHOD CALCPROFILE_10D0_A0LTAMAXT32T52 : BOOL
VAR_INPUT
	LRSTARTACC : LREAL;
	LRSTARTVEL : LREAL;
	LRMAXACC : LREAL;
	LRMAXVEL : LREAL;
	LRMAXDEC : LREAL;
	LRTARGETACC : LREAL;
	LRTARGETVEL : LREAL;
	LRTARGETPOS : LREAL;
	LRJERKTIMEACC : LREAL;
	LRJERKTIMEDEC : LREAL;
	LRJERKACC : LREAL;
	LRJERKDEC : LREAL;
END_VAR
VAR_IN_OUT
	SCPROFILEDATA : L_MB1P_ProfileData;
END_VAR
END_METHOD

METHOD CALCPROFILE_20A0 : BOOL
VAR_INPUT
	LRSTARTACC : LREAL;
	LRSTARTVEL : LREAL;
	LRMAXACC : LREAL;
	LRMAXDEC : LREAL;
	LRMAXVEL : LREAL;
	LRTARGETACC : LREAL;
	LRTARGETVEL : LREAL;
	LRTARGETPOS : LREAL;
	LRJERKACC : LREAL;
	LRJERKDEC : LREAL;
	LRJERKTIMEACC : LREAL;
	LRJERKTIMEDEC : LREAL;
END_VAR
VAR_OUTPUT
	DWSTATE : DWORD;
END_VAR
VAR_IN_OUT
	SCPROFILEDATA : L_MB1P_ProfileData;
	SCPROFILEPARAMETER : L_MB1P_ProfileParameter;
END_VAR
END_METHOD

METHOD CALCPROFILE_20A0_A0GTAMAXT71 : BOOL
VAR_INPUT
	LRSTARTACC : LREAL;
	LRSTARTVEL : LREAL;
	LRMAXACC : LREAL;
	LRMAXDEC : LREAL;
	LRMAXVEL : LREAL;
	LRTARGETACC : LREAL;
	LRTARGETVEL : LREAL;
	LRTARGETPOS : LREAL;
	LRJERKACC : LREAL;
	LRJERKDEC : LREAL;
	LRJERKTIMEACC : LREAL;
	LRJERKTIMEDEC : LREAL;
END_VAR
VAR_IN_OUT
	SCPROFILEDATA : L_MB1P_ProfileData;
END_VAR
END_METHOD

METHOD CALCPROFILE_20A0_A0GTAMAXT72 : BOOL
VAR_INPUT
	LRSTARTACC : LREAL;
	LRSTARTVEL : LREAL;
	LRMAXACC : LREAL;
	LRMAXDEC : LREAL;
	LRMAXVEL : LREAL;
	LRTARGETACC : LREAL;
	LRTARGETVEL : LREAL;
	LRTARGETPOS : LREAL;
	LRJERKACC : LREAL;
	LRJERKDEC : LREAL;
	LRJERKTIMEACC : LREAL;
	LRJERKTIMEDEC : LREAL;
END_VAR
VAR_IN_OUT
	SCPROFILEDATA : L_MB1P_ProfileData;
END_VAR
END_METHOD

METHOD CALCPROFILE_20A0_A0LTAMAXT71 : BOOL
VAR_INPUT
	LRSTARTACC : LREAL;
	LRSTARTVEL : LREAL;
	LRMAXACC : LREAL;
	LRMAXDEC : LREAL;
	LRMAXVEL : LREAL;
	LRTARGETACC : LREAL;
	LRTARGETVEL : LREAL;
	LRTARGETPOS : LREAL;
	LRJERKACC : LREAL;
	LRJERKDEC : LREAL;
	LRJERKTIMEACC : LREAL;
	LRJERKTIMEDEC : LREAL;
END_VAR
VAR_IN_OUT
	SCPROFILEDATA : L_MB1P_ProfileData;
END_VAR
END_METHOD

METHOD CALCPROFILE_20A0_A0LTAMAXT72 : BOOL
VAR_INPUT
	LRSTARTACC : LREAL;
	LRSTARTVEL : LREAL;
	LRMAXACC : LREAL;
	LRMAXDEC : LREAL;
	LRMAXVEL : LREAL;
	LRTARGETACC : LREAL;
	LRTARGETVEL : LREAL;
	LRTARGETPOS : LREAL;
	LRJERKACC : LREAL;
	LRJERKDEC : LREAL;
	LRJERKTIMEACC : LREAL;
	LRJERKTIMEDEC : LREAL;
END_VAR
VAR_IN_OUT
	SCPROFILEDATA : L_MB1P_ProfileData;
END_VAR
END_METHOD

METHOD CALCPROFILE_20B0 : BOOL
VAR_INPUT
	LRSTARTACC : LREAL;
	LRSTARTVEL : LREAL;
	LRMAXACC : LREAL;
	LRMAXDEC : LREAL;
	LRMAXVEL : LREAL;
	LRTARGETACC : LREAL;
	LRTARGETVEL : LREAL;
	LRTARGETPOS : LREAL;
	LRJERKACC : LREAL;
	LRJERKDEC : LREAL;
	LRJERKTIMEACC : LREAL;
	LRJERKTIMEDEC : LREAL;
	SCMAXPROFILEDATA : L_MB1P_IntProfileData;
	SCMINPROFILEDATA : L_MB1P_IntProfileData;
END_VAR
VAR_OUTPUT
	DWSTATE : DWORD;
END_VAR
VAR_IN_OUT
	SCPROFILEDATA : L_MB1P_ProfileData;
	SCPROFILEPARAMETER : L_MB1P_ProfileParameter;
END_VAR
END_METHOD

METHOD CALCPROFILE_20B0_A0GTAMAXSEARCHTIMEST5T7 : BOOL
VAR_INPUT
	LRSTARTACC : LREAL;
	LRSTARTVEL : LREAL;
	LRMAXACC : LREAL;
	LRMAXDEC : LREAL;
	LRMAXVEL : LREAL;
	LRTARGETACC : LREAL;
	LRTARGETVEL : LREAL;
	LRTARGETPOS : LREAL;
	LRJERKACC : LREAL;
	LRJERKDEC : LREAL;
	LRJERKTIMEACC : LREAL;
	LRJERKTIMEDEC : LREAL;
	T5_STARTVALUE : LREAL;
	T7_STARTVALUE : LREAL;
END_VAR
VAR_OUTPUT
	T5 : LREAL;
	T7 : LREAL;
END_VAR
END_METHOD

METHOD CALCPROFILE_20B0_A0GTAMAXT5T7 : BOOL
VAR_INPUT
	LRSTARTACC : LREAL;
	LRSTARTVEL : LREAL;
	LRMAXACC : LREAL;
	LRMAXDEC : LREAL;
	LRMAXVEL : LREAL;
	LRTARGETACC : LREAL;
	LRTARGETVEL : LREAL;
	LRTARGETPOS : LREAL;
	LRJERKACC : LREAL;
	LRJERKDEC : LREAL;
	LRJERKTIMEACC : LREAL;
	LRJERKTIMEDEC : LREAL;
	T5 : LREAL;
	T7 : LREAL;
END_VAR
VAR_IN_OUT
	SCPROFILEDATA : L_MB1P_ProfileData;
END_VAR
END_METHOD

METHOD CALCPROFILE_20B0_A0LTAMAXSEARCHTIMEST5T7 : BOOL
VAR_INPUT
	LRSTARTACC : LREAL;
	LRSTARTVEL : LREAL;
	LRMAXACC : LREAL;
	LRMAXDEC : LREAL;
	LRMAXVEL : LREAL;
	LRTARGETACC : LREAL;
	LRTARGETVEL : LREAL;
	LRTARGETPOS : LREAL;
	LRJERKACC : LREAL;
	LRJERKDEC : LREAL;
	LRJERKTIMEACC : LREAL;
	LRJERKTIMEDEC : LREAL;
	T5_STARTVALUE : LREAL;
	T7_STARTVALUE : LREAL;
END_VAR
VAR_OUTPUT
	T5 : LREAL;
	T7 : LREAL;
END_VAR
END_METHOD

METHOD CALCPROFILE_20B0_A0LTAMAXT5T7 : BOOL
VAR_INPUT
	LRSTARTACC : LREAL;
	LRSTARTVEL : LREAL;
	LRMAXACC : LREAL;
	LRMAXDEC : LREAL;
	LRMAXVEL : LREAL;
	LRTARGETACC : LREAL;
	LRTARGETVEL : LREAL;
	LRTARGETPOS : LREAL;
	LRJERKACC : LREAL;
	LRJERKDEC : LREAL;
	LRJERKTIMEACC : LREAL;
	LRJERKTIMEDEC : LREAL;
	T5 : LREAL;
	T7 : LREAL;
END_VAR
VAR_IN_OUT
	SCPROFILEDATA : L_MB1P_ProfileData;
END_VAR
END_METHOD

METHOD CALCPROFILE_20BA : BOOL
VAR_INPUT
	LRSTARTACC : LREAL;
	LRSTARTVEL : LREAL;
	LRMAXACC : LREAL;
	LRMAXDEC : LREAL;
	LRMAXVEL : LREAL;
	LRTARGETACC : LREAL;
	LRTARGETVEL : LREAL;
	LRTARGETPOS : LREAL;
	LRJERKACC : LREAL;
	LRJERKDEC : LREAL;
	LRJERKTIMEACC : LREAL;
	LRJERKTIMEDEC : LREAL;
	SCMAXPROFILEDATA : L_MB1P_IntProfileData;
	SCMINPROFILEDATA : L_MB1P_IntProfileData;
END_VAR
VAR_OUTPUT
	DWSTATE : DWORD;
END_VAR
VAR_IN_OUT
	SCPROFILEDATA : L_MB1P_ProfileData;
	SCPROFILEPARAMETER : L_MB1P_ProfileParameter;
END_VAR
END_METHOD

METHOD CALCPROFILE_20BA_A0GTAMAX : BOOL
VAR_INPUT
	LRSTARTACC : LREAL;
	LRSTARTVEL : LREAL;
	LRMAXACC : LREAL;
	LRMAXDEC : LREAL;
	LRMAXVEL : LREAL;
	LRTARGETACC : LREAL;
	LRTARGETVEL : LREAL;
	LRTARGETPOS : LREAL;
	LRJERKACC : LREAL;
	LRJERKDEC : LREAL;
	LRJERKTIMEACC : LREAL;
	LRJERKTIMEDEC : LREAL;
	T7 : LREAL;
END_VAR
VAR_IN_OUT
	SCPROFILEDATA : L_MB1P_ProfileData;
END_VAR
END_METHOD

METHOD CALCPROFILE_20BA_A0LETAMAX : BOOL
VAR_INPUT
	LRSTARTACC : LREAL;
	LRSTARTVEL : LREAL;
	LRMAXACC : LREAL;
	LRMAXDEC : LREAL;
	LRMAXVEL : LREAL;
	LRTARGETACC : LREAL;
	LRTARGETVEL : LREAL;
	LRTARGETPOS : LREAL;
	LRJERKACC : LREAL;
	LRJERKDEC : LREAL;
	LRJERKTIMEACC : LREAL;
	LRJERKTIMEDEC : LREAL;
	T7 : LREAL;
END_VAR
VAR_IN_OUT
	SCPROFILEDATA : L_MB1P_ProfileData;
END_VAR
END_METHOD

METHOD CALCPROFILE_20BA_AOGTAMAX_SEARCHTIMES : BOOL
VAR_INPUT
	LRSTARTACC : LREAL;
	LRSTARTVEL : LREAL;
	LRMAXACC : LREAL;
	LRMAXDEC : LREAL;
	LRMAXVEL : LREAL;
	LRTARGETACC : LREAL;
	LRTARGETVEL : LREAL;
	LRTARGETPOS : LREAL;
	LRJERKACC : LREAL;
	LRJERKDEC : LREAL;
	LRJERKTIMEACC : LREAL;
	LRJERKTIMEDEC : LREAL;
	T7_MINVALUE : LREAL;
	T7_MAXVALUE : LREAL;
END_VAR
VAR_OUTPUT
	T7 : LREAL;
END_VAR
END_METHOD

METHOD CALCPROFILE_20BA_AOLETAMAX_SEARCHTIMES : BOOL
VAR_INPUT
	LRSTARTACC : LREAL;
	LRSTARTVEL : LREAL;
	LRMAXACC : LREAL;
	LRMAXDEC : LREAL;
	LRMAXVEL : LREAL;
	LRTARGETACC : LREAL;
	LRTARGETVEL : LREAL;
	LRTARGETPOS : LREAL;
	LRJERKACC : LREAL;
	LRJERKDEC : LREAL;
	LRJERKTIMEACC : LREAL;
	LRJERKTIMEDEC : LREAL;
	T7_MINVALUE : LREAL;
	T7_MAXVALUE : LREAL;
END_VAR
VAR_OUTPUT
	T7 : LREAL;
END_VAR
END_METHOD

METHOD CALCPROFILE_20C0 : BOOL
VAR_INPUT
	LRSTARTACC : LREAL;
	LRSTARTVEL : LREAL;
	LRMAXACC : LREAL;
	LRMAXDEC : LREAL;
	LRMAXVEL : LREAL;
	LRTARGETACC : LREAL;
	LRTARGETVEL : LREAL;
	LRTARGETPOS : LREAL;
	LRJERKACC : LREAL;
	LRJERKDEC : LREAL;
	LRJERKTIMEACC : LREAL;
	LRJERKTIMEDEC : LREAL;
	SCMAXPROFILEDATA : L_MB1P_IntProfileData;
	SCMINPROFILEDATA : L_MB1P_IntProfileData;
END_VAR
VAR_OUTPUT
	DWSTATE : DWORD;
END_VAR
VAR_IN_OUT
	SCPROFILEDATA : L_MB1P_ProfileData;
	SCPROFILEPARAMETER : L_MB1P_ProfileParameter;
END_VAR
END_METHOD

METHOD CALCPROFILE_20C0_SEARCHTIMEST5T7 : BOOL
VAR_INPUT
	LRSTARTACC : LREAL;
	LRSTARTVEL : LREAL;
	LRMAXACC : LREAL;
	LRMAXDEC : LREAL;
	LRMAXVEL : LREAL;
	LRTARGETACC : LREAL;
	LRTARGETVEL : LREAL;
	LRTARGETPOS : LREAL;
	LRJERKACC : LREAL;
	LRJERKDEC : LREAL;
	LRJERKTIMEACC : LREAL;
	LRJERKTIMEDEC : LREAL;
	T5_STARTVALUE : LREAL;
	T7_STARTVALUE : LREAL;
END_VAR
VAR_OUTPUT
	T5 : LREAL;
	T7 : LREAL;
END_VAR
END_METHOD

METHOD CALCPROFILE_20C0_AELTAMAXT5T7 : BOOL
VAR_INPUT
	LRSTARTACC : LREAL;
	LRSTARTVEL : LREAL;
	LRMAXACC : LREAL;
	LRMAXDEC : LREAL;
	LRMAXVEL : LREAL;
	LRTARGETACC : LREAL;
	LRTARGETVEL : LREAL;
	LRTARGETPOS : LREAL;
	LRJERKACC : LREAL;
	LRJERKDEC : LREAL;
	LRJERKTIMEACC : LREAL;
	LRJERKTIMEDEC : LREAL;
	T5 : LREAL;
	T7 : LREAL;
END_VAR
VAR_IN_OUT
	SCPROFILEDATA : L_MB1P_ProfileData;
END_VAR
END_METHOD

METHOD CALCPROFILE_20CB : BOOL
VAR_INPUT
	LRSTARTACC : LREAL;
	LRSTARTVEL : LREAL;
	LRMAXACC : LREAL;
	LRMAXDEC : LREAL;
	LRMAXVEL : LREAL;
	LRTARGETACC : LREAL;
	LRTARGETVEL : LREAL;
	LRTARGETPOS : LREAL;
	LRJERKACC : LREAL;
	LRJERKDEC : LREAL;
	LRJERKTIMEACC : LREAL;
	LRJERKTIMEDEC : LREAL;
	SCMAXPROFILEDATA : L_MB1P_IntProfileData;
	SCMINPROFILEDATA : L_MB1P_IntProfileData;
END_VAR
VAR_OUTPUT
	DWSTATE : DWORD;
END_VAR
VAR_IN_OUT
	SCPROFILEDATA : L_MB1P_ProfileData;
	SCPROFILEPARAMETER : L_MB1P_ProfileParameter;
END_VAR
END_METHOD

METHOD CALCPROFILE_20CB_AOGET0 : BOOL
VAR_INPUT
	LRSTARTACC : LREAL;
	LRSTARTVEL : LREAL;
	LRMAXACC : LREAL;
	LRMAXDEC : LREAL;
	LRMAXVEL : LREAL;
	LRTARGETACC : LREAL;
	LRTARGETVEL : LREAL;
	LRTARGETPOS : LREAL;
	LRJERKACC : LREAL;
	LRJERKDEC : LREAL;
	LRJERKTIMEACC : LREAL;
	LRJERKTIMEDEC : LREAL;
	T7 : LREAL;
END_VAR
VAR_IN_OUT
	SCPROFILEDATA : L_MB1P_ProfileData;
END_VAR
END_METHOD

METHOD CALCPROFILE_20CB_AOLT0 : BOOL
VAR_INPUT
	LRSTARTACC : LREAL;
	LRSTARTVEL : LREAL;
	LRMAXACC : LREAL;
	LRMAXDEC : LREAL;
	LRMAXVEL : LREAL;
	LRTARGETACC : LREAL;
	LRTARGETVEL : LREAL;
	LRTARGETPOS : LREAL;
	LRJERKACC : LREAL;
	LRJERKDEC : LREAL;
	LRJERKTIMEACC : LREAL;
	LRJERKTIMEDEC : LREAL;
	T7 : LREAL;
END_VAR
VAR_IN_OUT
	SCPROFILEDATA : L_MB1P_ProfileData;
END_VAR
END_METHOD

METHOD CALCPROFILE_20CBAOGET0_SEARCHTIMES : BOOL
VAR_INPUT
	LRSTARTACC : LREAL;
	LRSTARTVEL : LREAL;
	LRMAXACC : LREAL;
	LRMAXDEC : LREAL;
	LRMAXVEL : LREAL;
	LRTARGETACC : LREAL;
	LRTARGETVEL : LREAL;
	LRTARGETPOS : LREAL;
	LRJERKACC : LREAL;
	LRJERKDEC : LREAL;
	LRJERKTIMEACC : LREAL;
	LRJERKTIMEDEC : LREAL;
	T7_MINVALUE : LREAL;
	T7_MAXVALUE : LREAL;
END_VAR
VAR_OUTPUT
	T7 : LREAL;
END_VAR
END_METHOD

METHOD CALCPROFILE_20CBAOLT0_SEARCHTIMES : BOOL
VAR_INPUT
	LRSTARTACC : LREAL;
	LRSTARTVEL : LREAL;
	LRMAXACC : LREAL;
	LRMAXDEC : LREAL;
	LRMAXVEL : LREAL;
	LRTARGETACC : LREAL;
	LRTARGETVEL : LREAL;
	LRTARGETPOS : LREAL;
	LRJERKACC : LREAL;
	LRJERKDEC : LREAL;
	LRJERKTIMEACC : LREAL;
	LRJERKTIMEDEC : LREAL;
	T7_MINVALUE : LREAL;
	T7_MAXVALUE : LREAL;
END_VAR
VAR_OUTPUT
	T7 : LREAL;
END_VAR
END_METHOD

METHOD CALCPROFILE_20D0 : BOOL
VAR_INPUT
	LRSTARTACC : LREAL;
	LRSTARTVEL : LREAL;
	LRMAXACC : LREAL;
	LRMAXDEC : LREAL;
	LRMAXVEL : LREAL;
	LRTARGETACC : LREAL;
	LRTARGETVEL : LREAL;
	LRTARGETPOS : LREAL;
	LRJERKACC : LREAL;
	LRJERKDEC : LREAL;
	LRJERKTIMEACC : LREAL;
	LRJERKTIMEDEC : LREAL;
	SCMAXPROFILEDATA : L_MB1P_IntProfileData;
	SCMINPROFILEDATA : L_MB1P_IntProfileData;
END_VAR
VAR_OUTPUT
	DWSTATE : DWORD;
END_VAR
VAR_IN_OUT
	SCPROFILEDATA : L_MB1P_ProfileData;
	SCPROFILEPARAMETER : L_MB1P_ProfileParameter;
END_VAR
END_METHOD

METHOD CALCPROFILE_20D0_SEARCHTIMEST5T7 : BOOL
VAR_INPUT
	LRSTARTACC : LREAL;
	LRSTARTVEL : LREAL;
	LRMAXACC : LREAL;
	LRMAXDEC : LREAL;
	LRMAXVEL : LREAL;
	LRTARGETACC : LREAL;
	LRTARGETVEL : LREAL;
	LRTARGETPOS : LREAL;
	LRJERKACC : LREAL;
	LRJERKDEC : LREAL;
	LRJERKTIMEACC : LREAL;
	LRJERKTIMEDEC : LREAL;
	T5_STARTVALUE : LREAL;
	T7_STARTVALUE : LREAL;
END_VAR
VAR_OUTPUT
	T5 : LREAL;
	T7 : LREAL;
END_VAR
END_METHOD

METHOD CALCPROFILE_20D0_A0LTAMAXT5T7 : BOOL
VAR_INPUT
	LRSTARTACC : LREAL;
	LRSTARTVEL : LREAL;
	LRMAXACC : LREAL;
	LRMAXDEC : LREAL;
	LRMAXVEL : LREAL;
	LRTARGETACC : LREAL;
	LRTARGETVEL : LREAL;
	LRTARGETPOS : LREAL;
	LRJERKACC : LREAL;
	LRJERKDEC : LREAL;
	LRJERKTIMEACC : LREAL;
	LRJERKTIMEDEC : LREAL;
	T5 : LREAL;
	T7 : LREAL;
END_VAR
VAR_IN_OUT
	SCPROFILEDATA : L_MB1P_ProfileData;
END_VAR
END_METHOD

METHOD CALCPROFILE_20D1 : BOOL
VAR_INPUT
	LRSTARTACC : LREAL;
	LRSTARTVEL : LREAL;
	LRMAXACC : LREAL;
	LRMAXDEC : LREAL;
	LRMAXVEL : LREAL;
	LRTARGETACC : LREAL;
	LRTARGETVEL : LREAL;
	LRTARGETPOS : LREAL;
	LRJERKACC : LREAL;
	LRJERKDEC : LREAL;
	LRJERKTIMEACC : LREAL;
	LRJERKTIMEDEC : LREAL;
	SCMAXPROFILEDATA : L_MB1P_IntProfileData;
	SCMINPROFILEDATA : L_MB1P_IntProfileData;
END_VAR
VAR_OUTPUT
	DWSTATE : DWORD;
END_VAR
VAR_IN_OUT
	SCPROFILEDATA : L_MB1P_ProfileData;
	SCPROFILEPARAMETER : L_MB1P_ProfileParameter;
END_VAR
END_METHOD

METHOD CALCPROFILE_20D1_AOGET0 : BOOL
VAR_INPUT
	LRSTARTACC : LREAL;
	LRSTARTVEL : LREAL;
	LRMAXACC : LREAL;
	LRMAXDEC : LREAL;
	LRMAXVEL : LREAL;
	LRTARGETACC : LREAL;
	LRTARGETVEL : LREAL;
	LRTARGETPOS : LREAL;
	LRJERKACC : LREAL;
	LRJERKDEC : LREAL;
	LRJERKTIMEACC : LREAL;
	LRJERKTIMEDEC : LREAL;
	T7 : LREAL;
END_VAR
VAR_IN_OUT
	SCPROFILEDATA : L_MB1P_ProfileData;
END_VAR
END_METHOD

METHOD CALCPROFILE_20D1_AOLT0 : BOOL
VAR_INPUT
	LRSTARTACC : LREAL;
	LRSTARTVEL : LREAL;
	LRMAXACC : LREAL;
	LRMAXDEC : LREAL;
	LRMAXVEL : LREAL;
	LRTARGETACC : LREAL;
	LRTARGETVEL : LREAL;
	LRTARGETPOS : LREAL;
	LRJERKACC : LREAL;
	LRJERKDEC : LREAL;
	LRJERKTIMEACC : LREAL;
	LRJERKTIMEDEC : LREAL;
	T7 : LREAL;
END_VAR
VAR_IN_OUT
	SCPROFILEDATA : L_MB1P_ProfileData;
END_VAR
END_METHOD

METHOD CALCPROFILE_20D1AOGET0_SEARCHTIMES : BOOL
VAR_INPUT
	LRSTARTACC : LREAL;
	LRSTARTVEL : LREAL;
	LRMAXACC : LREAL;
	LRMAXDEC : LREAL;
	LRMAXVEL : LREAL;
	LRTARGETACC : LREAL;
	LRTARGETVEL : LREAL;
	LRTARGETPOS : LREAL;
	LRJERKACC : LREAL;
	LRJERKDEC : LREAL;
	LRJERKTIMEACC : LREAL;
	LRJERKTIMEDEC : LREAL;
	T7_STARTVALUE : LREAL;
END_VAR
VAR_OUTPUT
	T7 : LREAL;
END_VAR
END_METHOD

METHOD CALCPROFILE_20D1AOLT0_SEARCHTIMES : BOOL
VAR_INPUT
	LRSTARTACC : LREAL;
	LRSTARTVEL : LREAL;
	LRMAXACC : LREAL;
	LRMAXDEC : LREAL;
	LRMAXVEL : LREAL;
	LRTARGETACC : LREAL;
	LRTARGETVEL : LREAL;
	LRTARGETPOS : LREAL;
	LRJERKACC : LREAL;
	LRJERKDEC : LREAL;
	LRJERKTIMEACC : LREAL;
	LRJERKTIMEDEC : LREAL;
	T7_STARTVALUE : LREAL;
END_VAR
VAR_OUTPUT
	T7 : LREAL;
END_VAR
END_METHOD

METHOD CALCPROFILE_20DA : BOOL
VAR_INPUT
	LRSTARTACC : LREAL;
	LRSTARTVEL : LREAL;
	LRMAXACC : LREAL;
	LRMAXDEC : LREAL;
	LRMAXVEL : LREAL;
	LRTARGETACC : LREAL;
	LRTARGETVEL : LREAL;
	LRTARGETPOS : LREAL;
	LRJERKACC : LREAL;
	LRJERKDEC : LREAL;
	LRJERKTIMEACC : LREAL;
	LRJERKTIMEDEC : LREAL;
	SCMAXPROFILEDATA : L_MB1P_IntProfileData;
	SCMINPROFILEDATA : L_MB1P_IntProfileData;
END_VAR
VAR_OUTPUT
	DWSTATE : DWORD;
END_VAR
VAR_IN_OUT
	SCPROFILEDATA : L_MB1P_ProfileData;
	SCPROFILEPARAMETER : L_MB1P_ProfileParameter;
END_VAR
END_METHOD

METHOD CALCPROFILE_20DA_AELT0 : BOOL
VAR_INPUT
	LRSTARTACC : LREAL;
	LRSTARTVEL : LREAL;
	LRMAXACC : LREAL;
	LRMAXDEC : LREAL;
	LRMAXVEL : LREAL;
	LRTARGETACC : LREAL;
	LRTARGETVEL : LREAL;
	LRTARGETPOS : LREAL;
	LRJERKACC : LREAL;
	LRJERKDEC : LREAL;
	LRJERKTIMEACC : LREAL;
	LRJERKTIMEDEC : LREAL;
	T7 : LREAL;
END_VAR
VAR_IN_OUT
	SCPROFILEDATA : L_MB1P_ProfileData;
END_VAR
END_METHOD

METHOD CALCPROFILE_20DAAELT0_SEARCHTIMES : BOOL
VAR_INPUT
	LRSTARTACC : LREAL;
	LRSTARTVEL : LREAL;
	LRMAXACC : LREAL;
	LRMAXDEC : LREAL;
	LRMAXVEL : LREAL;
	LRTARGETACC : LREAL;
	LRTARGETVEL : LREAL;
	LRTARGETPOS : LREAL;
	LRJERKACC : LREAL;
	LRJERKDEC : LREAL;
	LRJERKTIMEACC : LREAL;
	LRJERKTIMEDEC : LREAL;
	T7_MINVALUE : LREAL;
	T7_MAXVALUE : LREAL;
END_VAR
VAR_OUTPUT
	T7 : LREAL;
END_VAR
END_METHOD

METHOD CALCPROFILE_20DB : BOOL
VAR_INPUT
	LRSTARTACC : LREAL;
	LRSTARTVEL : LREAL;
	LRMAXACC : LREAL;
	LRMAXDEC : LREAL;
	LRMAXVEL : LREAL;
	LRTARGETACC : LREAL;
	LRTARGETVEL : LREAL;
	LRTARGETPOS : LREAL;
	LRJERKACC : LREAL;
	LRJERKDEC : LREAL;
	LRJERKTIMEACC : LREAL;
	LRJERKTIMEDEC : LREAL;
	SCMAXPROFILEDATA : L_MB1P_IntProfileData;
	SCMINPROFILEDATA : L_MB1P_IntProfileData;
END_VAR
VAR_OUTPUT
	DWSTATE : DWORD;
END_VAR
VAR_IN_OUT
	SCPROFILEDATA : L_MB1P_ProfileData;
	SCPROFILEPARAMETER : L_MB1P_ProfileParameter;
END_VAR
END_METHOD

METHOD CALCPROFILE_20DB_AOGET0 : BOOL
VAR_INPUT
	LRSTARTACC : LREAL;
	LRSTARTVEL : LREAL;
	LRMAXACC : LREAL;
	LRMAXDEC : LREAL;
	LRMAXVEL : LREAL;
	LRTARGETACC : LREAL;
	LRTARGETVEL : LREAL;
	LRTARGETPOS : LREAL;
	LRJERKACC : LREAL;
	LRJERKDEC : LREAL;
	LRJERKTIMEACC : LREAL;
	LRJERKTIMEDEC : LREAL;
	T7 : LREAL;
END_VAR
VAR_IN_OUT
	SCPROFILEDATA : L_MB1P_ProfileData;
END_VAR
END_METHOD

METHOD CALCPROFILE_20DB_AOLT0 : BOOL
VAR_INPUT
	LRSTARTACC : LREAL;
	LRSTARTVEL : LREAL;
	LRMAXACC : LREAL;
	LRMAXDEC : LREAL;
	LRMAXVEL : LREAL;
	LRTARGETACC : LREAL;
	LRTARGETVEL : LREAL;
	LRTARGETPOS : LREAL;
	LRJERKACC : LREAL;
	LRJERKDEC : LREAL;
	LRJERKTIMEACC : LREAL;
	LRJERKTIMEDEC : LREAL;
	T7 : LREAL;
END_VAR
VAR_IN_OUT
	SCPROFILEDATA : L_MB1P_ProfileData;
END_VAR
END_METHOD

METHOD CALCPROFILE_20DBAOGET0_SEARCHTIMES : BOOL
VAR_INPUT
	LRSTARTACC : LREAL;
	LRSTARTVEL : LREAL;
	LRMAXACC : LREAL;
	LRMAXDEC : LREAL;
	LRMAXVEL : LREAL;
	LRTARGETACC : LREAL;
	LRTARGETVEL : LREAL;
	LRTARGETPOS : LREAL;
	LRJERKACC : LREAL;
	LRJERKDEC : LREAL;
	LRJERKTIMEACC : LREAL;
	LRJERKTIMEDEC : LREAL;
	T7_MINVALUE : LREAL;
	T7_MAXVALUE : LREAL;
END_VAR
VAR_OUTPUT
	T7 : LREAL;
END_VAR
END_METHOD

METHOD CALCPROFILE_20DBAOLT0_SEARCHTIMES : BOOL
VAR_INPUT
	LRSTARTACC : LREAL;
	LRSTARTVEL : LREAL;
	LRMAXACC : LREAL;
	LRMAXDEC : LREAL;
	LRMAXVEL : LREAL;
	LRTARGETACC : LREAL;
	LRTARGETVEL : LREAL;
	LRTARGETPOS : LREAL;
	LRJERKACC : LREAL;
	LRJERKDEC : LREAL;
	LRJERKTIMEACC : LREAL;
	LRJERKTIMEDEC : LREAL;
	T7_MINVALUE : LREAL;
	T7_MAXVALUE : LREAL;
END_VAR
VAR_OUTPUT
	T7 : LREAL;
END_VAR
END_METHOD

METHOD CALCPROFILE_30A0 : BOOL
VAR_INPUT
	LRSTARTACC : LREAL;
	LRSTARTVEL : LREAL;
	LRMAXACC : LREAL;
	LRMAXDEC : LREAL;
	LRMAXVEL : LREAL;
	LRTARGETACC : LREAL;
	LRTARGETVEL : LREAL;
	LRTARGETPOS : LREAL;
	LRJERKACC : LREAL;
	LRJERKDEC : LREAL;
	LRJERKTIMEACC : LREAL;
	LRJERKTIMEDEC : LREAL;
END_VAR
VAR_OUTPUT
	DWSTATE : DWORD;
END_VAR
VAR_IN_OUT
	SCPROFILEDATA : L_MB1P_ProfileData;
	SCPROFILEPARAMETER : L_MB1P_ProfileParameter;
END_VAR
END_METHOD

METHOD CALCPROFILE_30A0_A0GTAMAX : BOOL
VAR_INPUT
	LRSTARTACC : LREAL;
	LRSTARTVEL : LREAL;
	LRMAXACC : LREAL;
	LRMAXDEC : LREAL;
	LRMAXVEL : LREAL;
	LRTARGETACC : LREAL;
	LRTARGETVEL : LREAL;
	LRTARGETPOS : LREAL;
	LRJERKACC : LREAL;
	LRJERKDEC : LREAL;
	LRJERKTIMEACC : LREAL;
	LRJERKTIMEDEC : LREAL;
END_VAR
VAR_IN_OUT
	SCPROFILEDATA : L_MB1P_ProfileData;
END_VAR
END_METHOD

METHOD CALCPROFILE_30A0_A0LTAMAX : BOOL
VAR_INPUT
	LRSTARTACC : LREAL;
	LRSTARTVEL : LREAL;
	LRMAXACC : LREAL;
	LRMAXDEC : LREAL;
	LRMAXVEL : LREAL;
	LRTARGETACC : LREAL;
	LRTARGETVEL : LREAL;
	LRTARGETPOS : LREAL;
	LRJERKACC : LREAL;
	LRJERKDEC : LREAL;
	LRJERKTIMEACC : LREAL;
	LRJERKTIMEDEC : LREAL;
END_VAR
VAR_IN_OUT
	SCPROFILEDATA : L_MB1P_ProfileData;
END_VAR
END_METHOD

METHOD CALCPROFILE_30B0 : BOOL
VAR_INPUT
	LRSTARTACC : LREAL;
	LRSTARTVEL : LREAL;
	LRMAXACC : LREAL;
	LRMAXDEC : LREAL;
	LRMAXVEL : LREAL;
	LRTARGETACC : LREAL;
	LRTARGETVEL : LREAL;
	LRTARGETPOS : LREAL;
	LRJERKACC : LREAL;
	LRJERKDEC : LREAL;
	LRJERKTIMEACC : LREAL;
	LRJERKTIMEDEC : LREAL;
END_VAR
VAR_OUTPUT
	DWSTATE : DWORD;
END_VAR
VAR_IN_OUT
	SCPROFILEDATA : L_MB1P_ProfileData;
	SCPROFILEPARAMETER : L_MB1P_ProfileParameter;
END_VAR
END_METHOD

METHOD CALCPROFILE_30B0_A0GTAMAXT51 : BOOL
VAR_INPUT
	LRSTARTACC : LREAL;
	LRSTARTVEL : LREAL;
	LRMAXACC : LREAL;
	LRMAXDEC : LREAL;
	LRMAXVEL : LREAL;
	LRTARGETACC : LREAL;
	LRTARGETVEL : LREAL;
	LRTARGETPOS : LREAL;
	LRJERKACC : LREAL;
	LRJERKDEC : LREAL;
	LRJERKTIMEACC : LREAL;
	LRJERKTIMEDEC : LREAL;
END_VAR
VAR_IN_OUT
	SCPROFILEDATA : L_MB1P_ProfileData;
END_VAR
END_METHOD

METHOD CALCPROFILE_30B0_A0GTAMAXT52 : BOOL
VAR_INPUT
	LRSTARTACC : LREAL;
	LRSTARTVEL : LREAL;
	LRMAXACC : LREAL;
	LRMAXDEC : LREAL;
	LRMAXVEL : LREAL;
	LRTARGETACC : LREAL;
	LRTARGETVEL : LREAL;
	LRTARGETPOS : LREAL;
	LRJERKACC : LREAL;
	LRJERKDEC : LREAL;
	LRJERKTIMEACC : LREAL;
	LRJERKTIMEDEC : LREAL;
END_VAR
VAR_IN_OUT
	SCPROFILEDATA : L_MB1P_ProfileData;
END_VAR
END_METHOD

METHOD CALCPROFILE_30B0_A0LTAMAXT51 : BOOL
VAR_INPUT
	LRSTARTACC : LREAL;
	LRSTARTVEL : LREAL;
	LRMAXACC : LREAL;
	LRMAXDEC : LREAL;
	LRMAXVEL : LREAL;
	LRTARGETACC : LREAL;
	LRTARGETVEL : LREAL;
	LRTARGETPOS : LREAL;
	LRJERKACC : LREAL;
	LRJERKDEC : LREAL;
	LRJERKTIMEACC : LREAL;
	LRJERKTIMEDEC : LREAL;
END_VAR
VAR_IN_OUT
	SCPROFILEDATA : L_MB1P_ProfileData;
END_VAR
END_METHOD

METHOD CALCPROFILE_30B0_A0LTAMAXT52 : BOOL
VAR_INPUT
	LRSTARTACC : LREAL;
	LRSTARTVEL : LREAL;
	LRMAXACC : LREAL;
	LRMAXDEC : LREAL;
	LRMAXVEL : LREAL;
	LRTARGETACC : LREAL;
	LRTARGETVEL : LREAL;
	LRTARGETPOS : LREAL;
	LRJERKACC : LREAL;
	LRJERKDEC : LREAL;
	LRJERKTIMEACC : LREAL;
	LRJERKTIMEDEC : LREAL;
END_VAR
VAR_IN_OUT
	SCPROFILEDATA : L_MB1P_ProfileData;
END_VAR
END_METHOD

METHOD CALCPROFILE_30C0 : BOOL
VAR_INPUT
	LRSTARTACC : LREAL;
	LRSTARTVEL : LREAL;
	LRMAXACC : LREAL;
	LRMAXDEC : LREAL;
	LRMAXVEL : LREAL;
	LRTARGETACC : LREAL;
	LRTARGETVEL : LREAL;
	LRTARGETPOS : LREAL;
	LRJERKACC : LREAL;
	LRJERKDEC : LREAL;
	LRJERKTIMEACC : LREAL;
	LRJERKTIMEDEC : LREAL;
END_VAR
VAR_OUTPUT
	DWSTATE : DWORD;
END_VAR
VAR_IN_OUT
	SCPROFILEDATA : L_MB1P_ProfileData;
	SCPROFILEPARAMETER : L_MB1P_ProfileParameter;
END_VAR
END_METHOD

METHOD CALCPROFILE_30C0_A0GTAMAXT31 : BOOL
VAR_INPUT
	LRSTARTACC : LREAL;
	LRSTARTVEL : LREAL;
	LRMAXACC : LREAL;
	LRMAXDEC : LREAL;
	LRMAXVEL : LREAL;
	LRTARGETACC : LREAL;
	LRTARGETVEL : LREAL;
	LRTARGETPOS : LREAL;
	LRJERKACC : LREAL;
	LRJERKDEC : LREAL;
	LRJERKTIMEACC : LREAL;
	LRJERKTIMEDEC : LREAL;
END_VAR
VAR_IN_OUT
	SCPROFILEDATA : L_MB1P_ProfileData;
END_VAR
END_METHOD

METHOD CALCPROFILE_30C0_A0GTAMAXT32 : BOOL
VAR_INPUT
	LRSTARTACC : LREAL;
	LRSTARTVEL : LREAL;
	LRMAXACC : LREAL;
	LRMAXDEC : LREAL;
	LRMAXVEL : LREAL;
	LRTARGETACC : LREAL;
	LRTARGETVEL : LREAL;
	LRTARGETPOS : LREAL;
	LRJERKACC : LREAL;
	LRJERKDEC : LREAL;
	LRJERKTIMEACC : LREAL;
	LRJERKTIMEDEC : LREAL;
END_VAR
VAR_IN_OUT
	SCPROFILEDATA : L_MB1P_ProfileData;
END_VAR
END_METHOD

METHOD CALCPROFILE_30CB : BOOL
VAR_INPUT
	LRSTARTACC : LREAL;
	LRSTARTVEL : LREAL;
	LRMAXACC : LREAL;
	LRMAXDEC : LREAL;
	LRMAXVEL : LREAL;
	LRTARGETACC : LREAL;
	LRTARGETVEL : LREAL;
	LRTARGETPOS : LREAL;
	LRJERKACC : LREAL;
	LRJERKDEC : LREAL;
	LRJERKTIMEACC : LREAL;
	LRJERKTIMEDEC : LREAL;
	SCMAXPROFILEDATA : L_MB1P_IntProfileData;
	SCMINPROFILEDATA : L_MB1P_IntProfileData;
END_VAR
VAR_OUTPUT
	DWSTATE : DWORD;
END_VAR
VAR_IN_OUT
	SCPROFILEDATA : L_MB1P_ProfileData;
	SCPROFILEPARAMETER : L_MB1P_ProfileParameter;
END_VAR
END_METHOD

METHOD CALCPROFILE_30CB_PROFILEDATA : BOOL
VAR_INPUT
	LRSTARTACC : LREAL;
	LRSTARTVEL : LREAL;
	LRMAXACC : LREAL;
	LRMAXDEC : LREAL;
	LRMAXVEL : LREAL;
	LRTARGETACC : LREAL;
	LRTARGETVEL : LREAL;
	LRTARGETPOS : LREAL;
	LRJERKACC : LREAL;
	LRJERKDEC : LREAL;
	LRJERKTIMEACC : LREAL;
	LRJERKTIMEDEC : LREAL;
	T7 : LREAL;
END_VAR
VAR_IN_OUT
	SCPROFILEDATA : L_MB1P_ProfileData;
END_VAR
END_METHOD

METHOD CALCPROFILE_30CB_SEARCHTIMES : BOOL
VAR_INPUT
	LRSTARTACC : LREAL;
	LRSTARTVEL : LREAL;
	LRMAXACC : LREAL;
	LRMAXDEC : LREAL;
	LRMAXVEL : LREAL;
	LRTARGETACC : LREAL;
	LRTARGETVEL : LREAL;
	LRTARGETPOS : LREAL;
	LRJERKACC : LREAL;
	LRJERKDEC : LREAL;
	LRJERKTIMEACC : LREAL;
	LRJERKTIMEDEC : LREAL;
	T7_MINVALUE : LREAL;
	T7_MAXVALUE : LREAL;
END_VAR
VAR_OUTPUT
	T7 : LREAL;
END_VAR
END_METHOD

METHOD CALCPROFILE_30D0 : BOOL
VAR_INPUT
	LRSTARTACC : LREAL;
	LRSTARTVEL : LREAL;
	LRMAXACC : LREAL;
	LRMAXDEC : LREAL;
	LRMAXVEL : LREAL;
	LRTARGETACC : LREAL;
	LRTARGETVEL : LREAL;
	LRTARGETPOS : LREAL;
	LRJERKACC : LREAL;
	LRJERKDEC : LREAL;
	LRJERKTIMEACC : LREAL;
	LRJERKTIMEDEC : LREAL;
END_VAR
VAR_OUTPUT
	DWSTATE : DWORD;
END_VAR
VAR_IN_OUT
	SCPROFILEDATA : L_MB1P_ProfileData;
	SCPROFILEPARAMETER : L_MB1P_ProfileParameter;
END_VAR
END_METHOD

METHOD CALCPROFILE_30D0_A0GTAMAXT31T51 : BOOL
VAR_INPUT
	LRSTARTACC : LREAL;
	LRSTARTVEL : LREAL;
	LRMAXACC : LREAL;
	LRMAXDEC : LREAL;
	LRMAXVEL : LREAL;
	LRTARGETACC : LREAL;
	LRTARGETVEL : LREAL;
	LRTARGETPOS : LREAL;
	LRJERKACC : LREAL;
	LRJERKDEC : LREAL;
	LRJERKTIMEACC : LREAL;
	LRJERKTIMEDEC : LREAL;
END_VAR
VAR_IN_OUT
	SCPROFILEDATA : L_MB1P_ProfileData;
END_VAR
END_METHOD

METHOD CALCPROFILE_30D0_A0GTAMAXT31T52 : BOOL
VAR_INPUT
	LRSTARTACC : LREAL;
	LRSTARTVEL : LREAL;
	LRMAXACC : LREAL;
	LRMAXDEC : LREAL;
	LRMAXVEL : LREAL;
	LRTARGETACC : LREAL;
	LRTARGETVEL : LREAL;
	LRTARGETPOS : LREAL;
	LRJERKACC : LREAL;
	LRJERKDEC : LREAL;
	LRJERKTIMEACC : LREAL;
	LRJERKTIMEDEC : LREAL;
END_VAR
VAR_IN_OUT
	SCPROFILEDATA : L_MB1P_ProfileData;
END_VAR
END_METHOD

METHOD CALCPROFILE_30D0_A0GTAMAXT32T51 : BOOL
VAR_INPUT
	LRSTARTACC : LREAL;
	LRSTARTVEL : LREAL;
	LRMAXACC : LREAL;
	LRMAXDEC : LREAL;
	LRMAXVEL : LREAL;
	LRTARGETACC : LREAL;
	LRTARGETVEL : LREAL;
	LRTARGETPOS : LREAL;
	LRJERKACC : LREAL;
	LRJERKDEC : LREAL;
	LRJERKTIMEACC : LREAL;
	LRJERKTIMEDEC : LREAL;
END_VAR
VAR_IN_OUT
	SCPROFILEDATA : L_MB1P_ProfileData;
END_VAR
END_METHOD

METHOD CALCPROFILE_30D0_A0GTAMAXT32T52 : BOOL
VAR_INPUT
	LRSTARTACC : LREAL;
	LRSTARTVEL : LREAL;
	LRMAXACC : LREAL;
	LRMAXDEC : LREAL;
	LRMAXVEL : LREAL;
	LRTARGETACC : LREAL;
	LRTARGETVEL : LREAL;
	LRTARGETPOS : LREAL;
	LRJERKACC : LREAL;
	LRJERKDEC : LREAL;
	LRJERKTIMEACC : LREAL;
	LRJERKTIMEDEC : LREAL;
END_VAR
VAR_IN_OUT
	SCPROFILEDATA : L_MB1P_ProfileData;
END_VAR
END_METHOD

METHOD CALCPROFILE_30D1 : BOOL
VAR_INPUT
	LRSTARTACC : LREAL;
	LRSTARTVEL : LREAL;
	LRMAXACC : LREAL;
	LRMAXDEC : LREAL;
	LRMAXVEL : LREAL;
	LRTARGETACC : LREAL;
	LRTARGETVEL : LREAL;
	LRTARGETPOS : LREAL;
	LRJERKACC : LREAL;
	LRJERKDEC : LREAL;
	LRJERKTIMEACC : LREAL;
	LRJERKTIMEDEC : LREAL;
	SCMAXPROFILEDATA : L_MB1P_IntProfileData;
	SCMINPROFILEDATA : L_MB1P_IntProfileData;
END_VAR
VAR_OUTPUT
	DWSTATE : DWORD;
END_VAR
VAR_IN_OUT
	SCPROFILEDATA : L_MB1P_ProfileData;
	SCPROFILEPARAMETER : L_MB1P_ProfileParameter;
END_VAR
END_METHOD

METHOD CALCPROFILE_30D1_PROFILEDATA : BOOL
VAR_INPUT
	LRSTARTACC : LREAL;
	LRSTARTVEL : LREAL;
	LRMAXACC : LREAL;
	LRMAXDEC : LREAL;
	LRMAXVEL : LREAL;
	LRTARGETACC : LREAL;
	LRTARGETVEL : LREAL;
	LRTARGETPOS : LREAL;
	LRJERKACC : LREAL;
	LRJERKDEC : LREAL;
	LRJERKTIMEACC : LREAL;
	LRJERKTIMEDEC : LREAL;
	T7 : LREAL;
END_VAR
VAR_IN_OUT
	SCPROFILEDATA : L_MB1P_ProfileData;
END_VAR
END_METHOD

METHOD CALCPROFILE_30D1_SEARCHTIMES : BOOL
VAR_INPUT
	LRSTARTACC : LREAL;
	LRSTARTVEL : LREAL;
	LRMAXACC : LREAL;
	LRMAXDEC : LREAL;
	LRMAXVEL : LREAL;
	LRTARGETACC : LREAL;
	LRTARGETVEL : LREAL;
	LRTARGETPOS : LREAL;
	LRJERKACC : LREAL;
	LRJERKDEC : LREAL;
	LRJERKTIMEACC : LREAL;
	LRJERKTIMEDEC : LREAL;
	T7_MINVALUE : LREAL;
	T7_MAXVALUE : LREAL;
END_VAR
VAR_OUTPUT
	T7 : LREAL;
END_VAR
END_METHOD

METHOD CALCPROFILE_30DB : BOOL
VAR_INPUT
	LRSTARTACC : LREAL;
	LRSTARTVEL : LREAL;
	LRMAXACC : LREAL;
	LRMAXDEC : LREAL;
	LRMAXVEL : LREAL;
	LRTARGETACC : LREAL;
	LRTARGETVEL : LREAL;
	LRTARGETPOS : LREAL;
	LRJERKACC : LREAL;
	LRJERKDEC : LREAL;
	LRJERKTIMEACC : LREAL;
	LRJERKTIMEDEC : LREAL;
	SCMAXPROFILEDATA : L_MB1P_IntProfileData;
	SCMINPROFILEDATA : L_MB1P_IntProfileData;
END_VAR
VAR_OUTPUT
	DWSTATE : DWORD;
END_VAR
VAR_IN_OUT
	SCPROFILEDATA : L_MB1P_ProfileData;
	SCPROFILEPARAMETER : L_MB1P_ProfileParameter;
END_VAR
END_METHOD

METHOD CALCPROFILE_30DB_PROFILEDATA : BOOL
VAR_INPUT
	LRSTARTACC : LREAL;
	LRSTARTVEL : LREAL;
	LRMAXACC : LREAL;
	LRMAXDEC : LREAL;
	LRMAXVEL : LREAL;
	LRTARGETACC : LREAL;
	LRTARGETVEL : LREAL;
	LRTARGETPOS : LREAL;
	LRJERKACC : LREAL;
	LRJERKDEC : LREAL;
	LRJERKTIMEACC : LREAL;
	LRJERKTIMEDEC : LREAL;
	T7 : LREAL;
END_VAR
VAR_IN_OUT
	SCPROFILEDATA : L_MB1P_ProfileData;
END_VAR
END_METHOD

METHOD CALCPROFILE_30DB_SEARCHTIMES : BOOL
VAR_INPUT
	LRSTARTACC : LREAL;
	LRSTARTVEL : LREAL;
	LRMAXACC : LREAL;
	LRMAXDEC : LREAL;
	LRMAXVEL : LREAL;
	LRTARGETACC : LREAL;
	LRTARGETVEL : LREAL;
	LRTARGETPOS : LREAL;
	LRJERKACC : LREAL;
	LRJERKDEC : LREAL;
	LRJERKTIMEACC : LREAL;
	LRJERKTIMEDEC : LREAL;
	T7_MINVALUE : LREAL;
	T7_MAXVALUE : LREAL;
END_VAR
VAR_OUTPUT
	T7 : LREAL;
END_VAR
END_METHOD

METHOD CALCPROFILE_40A0 : BOOL
VAR_INPUT
	LRSTARTACC : LREAL;
	LRSTARTVEL : LREAL;
	LRMAXACC : LREAL;
	LRMAXDEC : LREAL;
	LRMAXVEL : LREAL;
	LRTARGETACC : LREAL;
	LRTARGETVEL : LREAL;
	LRTARGETPOS : LREAL;
	LRJERKACC : LREAL;
	LRJERKDEC : LREAL;
	LRJERKTIMEACC : LREAL;
	LRJERKTIMEDEC : LREAL;
END_VAR
VAR_OUTPUT
	DWSTATE : DWORD;
END_VAR
VAR_IN_OUT
	SCPROFILEDATA : L_MB1P_ProfileData;
	SCPROFILEPARAMETER : L_MB1P_ProfileParameter;
END_VAR
END_METHOD

METHOD CALCPROFILE_40A0_A0GTAMAX : BOOL
VAR_INPUT
	LRSTARTACC : LREAL;
	LRSTARTVEL : LREAL;
	LRMAXACC : LREAL;
	LRMAXDEC : LREAL;
	LRMAXVEL : LREAL;
	LRTARGETACC : LREAL;
	LRTARGETVEL : LREAL;
	LRTARGETPOS : LREAL;
	LRJERKACC : LREAL;
	LRJERKDEC : LREAL;
	LRJERKTIMEACC : LREAL;
	LRJERKTIMEDEC : LREAL;
END_VAR
VAR_IN_OUT
	SCPROFILEDATA : L_MB1P_ProfileData;
END_VAR
END_METHOD

METHOD CALCPROFILE_40A0_A0LTAMAX : BOOL
VAR_INPUT
	LRSTARTACC : LREAL;
	LRSTARTVEL : LREAL;
	LRMAXACC : LREAL;
	LRMAXDEC : LREAL;
	LRMAXVEL : LREAL;
	LRTARGETACC : LREAL;
	LRTARGETVEL : LREAL;
	LRTARGETPOS : LREAL;
	LRJERKACC : LREAL;
	LRJERKDEC : LREAL;
	LRJERKTIMEACC : LREAL;
	LRJERKTIMEDEC : LREAL;
END_VAR
VAR_IN_OUT
	SCPROFILEDATA : L_MB1P_ProfileData;
END_VAR
END_METHOD

METHOD CALCPROFILE_40B0 : BOOL
VAR_INPUT
	LRSTARTACC : LREAL;
	LRSTARTVEL : LREAL;
	LRMAXACC : LREAL;
	LRMAXDEC : LREAL;
	LRMAXVEL : LREAL;
	LRTARGETACC : LREAL;
	LRTARGETVEL : LREAL;
	LRTARGETPOS : LREAL;
	LRJERKACC : LREAL;
	LRJERKDEC : LREAL;
	LRJERKTIMEACC : LREAL;
	LRJERKTIMEDEC : LREAL;
END_VAR
VAR_OUTPUT
	DWSTATE : DWORD;
END_VAR
VAR_IN_OUT
	SCPROFILEDATA : L_MB1P_ProfileData;
	SCPROFILEPARAMETER : L_MB1P_ProfileParameter;
END_VAR
END_METHOD

METHOD CALCPROFILE_40C0 : BOOL
VAR_INPUT
	LRSTARTACC : LREAL;
	LRSTARTVEL : LREAL;
	LRMAXACC : LREAL;
	LRMAXDEC : LREAL;
	LRMAXVEL : LREAL;
	LRTARGETACC : LREAL;
	LRTARGETVEL : LREAL;
	LRTARGETPOS : LREAL;
	LRJERKACC : LREAL;
	LRJERKDEC : LREAL;
	LRJERKTIMEACC : LREAL;
	LRJERKTIMEDEC : LREAL;
END_VAR
VAR_OUTPUT
	DWSTATE : DWORD;
END_VAR
VAR_IN_OUT
	SCPROFILEDATA : L_MB1P_ProfileData;
	SCPROFILEPARAMETER : L_MB1P_ProfileParameter;
END_VAR
END_METHOD

METHOD CALCPROFILE_40C0_A0LTAMAXT31 : BOOL
VAR_INPUT
	LRSTARTACC : LREAL;
	LRSTARTVEL : LREAL;
	LRMAXACC : LREAL;
	LRMAXDEC : LREAL;
	LRMAXVEL : LREAL;
	LRTARGETACC : LREAL;
	LRTARGETVEL : LREAL;
	LRTARGETPOS : LREAL;
	LRJERKACC : LREAL;
	LRJERKDEC : LREAL;
	LRJERKTIMEACC : LREAL;
	LRJERKTIMEDEC : LREAL;
END_VAR
VAR_IN_OUT
	SCPROFILEDATA : L_MB1P_ProfileData;
END_VAR
END_METHOD

METHOD CALCPROFILE_40C0_A0LTAMAXT32 : BOOL
VAR_INPUT
	LRSTARTACC : LREAL;
	LRSTARTVEL : LREAL;
	LRMAXACC : LREAL;
	LRMAXDEC : LREAL;
	LRMAXVEL : LREAL;
	LRTARGETACC : LREAL;
	LRTARGETVEL : LREAL;
	LRTARGETPOS : LREAL;
	LRJERKACC : LREAL;
	LRJERKDEC : LREAL;
	LRJERKTIMEACC : LREAL;
	LRJERKTIMEDEC : LREAL;
END_VAR
VAR_IN_OUT
	SCPROFILEDATA : L_MB1P_ProfileData;
END_VAR
END_METHOD

METHOD CALCPROFILE_40D0 : BOOL
VAR_INPUT
	LRSTARTACC : LREAL;
	LRSTARTVEL : LREAL;
	LRMAXACC : LREAL;
	LRMAXDEC : LREAL;
	LRMAXVEL : LREAL;
	LRTARGETACC : LREAL;
	LRTARGETVEL : LREAL;
	LRTARGETPOS : LREAL;
	LRJERKACC : LREAL;
	LRJERKDEC : LREAL;
	LRJERKTIMEACC : LREAL;
	LRJERKTIMEDEC : LREAL;
END_VAR
VAR_OUTPUT
	DWSTATE : DWORD;
END_VAR
VAR_IN_OUT
	SCPROFILEDATA : L_MB1P_ProfileData;
	SCPROFILEPARAMETER : L_MB1P_ProfileParameter;
END_VAR
END_METHOD

METHOD CALCPROFILE_40E0 : BOOL
VAR_INPUT
	LRSTARTACC : LREAL;
	LRSTARTVEL : LREAL;
	LRMAXACC : LREAL;
	LRMAXDEC : LREAL;
	LRMAXVEL : LREAL;
	LRTARGETACC : LREAL;
	LRTARGETVEL : LREAL;
	LRTARGETPOS : LREAL;
	LRJERKACC : LREAL;
	LRJERKDEC : LREAL;
	LRJERKTIMEACC : LREAL;
	LRJERKTIMEDEC : LREAL;
END_VAR
VAR_OUTPUT
	DWSTATE : DWORD;
END_VAR
VAR_IN_OUT
	SCPROFILEDATA : L_MB1P_ProfileData;
	SCPROFILEPARAMETER : L_MB1P_ProfileParameter;
END_VAR
END_METHOD

METHOD CALCPROFILE_40F0 : BOOL
VAR_INPUT
	LRSTARTACC : LREAL;
	LRSTARTVEL : LREAL;
	LRMAXACC : LREAL;
	LRMAXDEC : LREAL;
	LRMAXVEL : LREAL;
	LRTARGETACC : LREAL;
	LRTARGETVEL : LREAL;
	LRTARGETPOS : LREAL;
	LRJERKACC : LREAL;
	LRJERKDEC : LREAL;
	LRJERKTIMEACC : LREAL;
	LRJERKTIMEDEC : LREAL;
END_VAR
VAR_OUTPUT
	DWSTATE : DWORD;
END_VAR
VAR_IN_OUT
	SCPROFILEDATA : L_MB1P_ProfileData;
	SCPROFILEPARAMETER : L_MB1P_ProfileParameter;
END_VAR
END_METHOD

METHOD CALCPROFILE_40F0_T51 : BOOL
VAR_INPUT
	LRSTARTACC : LREAL;
	LRSTARTVEL : LREAL;
	LRMAXACC : LREAL;
	LRMAXDEC : LREAL;
	LRMAXVEL : LREAL;
	LRTARGETACC : LREAL;
	LRTARGETVEL : LREAL;
	LRTARGETPOS : LREAL;
	LRJERKACC : LREAL;
	LRJERKDEC : LREAL;
	LRJERKTIMEACC : LREAL;
	LRJERKTIMEDEC : LREAL;
END_VAR
VAR_IN_OUT
	SCPROFILEDATA : L_MB1P_ProfileData;
END_VAR
END_METHOD

METHOD CALCPROFILE_40F0_T52 : BOOL
VAR_INPUT
	LRSTARTACC : LREAL;
	LRSTARTVEL : LREAL;
	LRMAXACC : LREAL;
	LRMAXDEC : LREAL;
	LRMAXVEL : LREAL;
	LRTARGETACC : LREAL;
	LRTARGETVEL : LREAL;
	LRTARGETPOS : LREAL;
	LRJERKACC : LREAL;
	LRJERKDEC : LREAL;
	LRJERKTIMEACC : LREAL;
	LRJERKTIMEDEC : LREAL;
END_VAR
VAR_IN_OUT
	SCPROFILEDATA : L_MB1P_ProfileData;
END_VAR
END_METHOD

METHOD CALCPROFILE_50A0 : BOOL
VAR_INPUT
	LRSTARTACC : LREAL;
	LRSTARTVEL : LREAL;
	LRMAXACC : LREAL;
	LRMAXDEC : LREAL;
	LRMAXVEL : LREAL;
	LRTARGETACC : LREAL;
	LRTARGETVEL : LREAL;
	LRTARGETPOS : LREAL;
	LRJERKACC : LREAL;
	LRJERKDEC : LREAL;
	LRJERKTIMEACC : LREAL;
	LRJERKTIMEDEC : LREAL;
END_VAR
VAR_OUTPUT
	DWSTATE : DWORD;
END_VAR
VAR_IN_OUT
	SCPROFILEDATA : L_MB1P_ProfileData;
	SCPROFILEPARAMETER : L_MB1P_ProfileParameter;
END_VAR
END_METHOD

METHOD CALCPROFILE_60A0 : BOOL
VAR_INPUT
	LRSTARTACC : LREAL;
	LRSTARTVEL : LREAL;
	LRMAXACC : LREAL;
	LRMAXDEC : LREAL;
	LRMAXVEL : LREAL;
	LRTARGETACC : LREAL;
	LRTARGETVEL : LREAL;
	LRTARGETPOS : LREAL;
	LRJERKACC : LREAL;
	LRJERKDEC : LREAL;
	LRJERKTIMEACC : LREAL;
	LRJERKTIMEDEC : LREAL;
END_VAR
VAR_OUTPUT
	DWSTATE : DWORD;
END_VAR
VAR_IN_OUT
	SCPROFILEDATA : L_MB1P_ProfileData;
	SCPROFILEPARAMETER : L_MB1P_ProfileParameter;
END_VAR
END_METHOD

METHOD CALCPROFILE_60A0_A0GTAMAX : BOOL
VAR_INPUT
	LRSTARTACC : LREAL;
	LRSTARTVEL : LREAL;
	LRMAXACC : LREAL;
	LRMAXDEC : LREAL;
	LRMAXVEL : LREAL;
	LRTARGETACC : LREAL;
	LRTARGETVEL : LREAL;
	LRTARGETPOS : LREAL;
	LRJERKACC : LREAL;
	LRJERKDEC : LREAL;
	LRJERKTIMEACC : LREAL;
	LRJERKTIMEDEC : LREAL;
END_VAR
VAR_IN_OUT
	SCPROFILEDATA : L_MB1P_ProfileData;
END_VAR
END_METHOD

METHOD CALCPROFILE_60A0_A0LTAMAX : BOOL
VAR_INPUT
	LRSTARTACC : LREAL;
	LRSTARTVEL : LREAL;
	LRMAXACC : LREAL;
	LRMAXDEC : LREAL;
	LRMAXVEL : LREAL;
	LRTARGETACC : LREAL;
	LRTARGETVEL : LREAL;
	LRTARGETPOS : LREAL;
	LRJERKACC : LREAL;
	LRJERKDEC : LREAL;
	LRJERKTIMEACC : LREAL;
	LRJERKTIMEDEC : LREAL;
END_VAR
VAR_IN_OUT
	SCPROFILEDATA : L_MB1P_ProfileData;
END_VAR
END_METHOD

METHOD CALCPROFILE_60B0 : BOOL
VAR_INPUT
	LRSTARTACC : LREAL;
	LRSTARTVEL : LREAL;
	LRMAXACC : LREAL;
	LRMAXDEC : LREAL;
	LRMAXVEL : LREAL;
	LRTARGETACC : LREAL;
	LRTARGETVEL : LREAL;
	LRTARGETPOS : LREAL;
	LRJERKACC : LREAL;
	LRJERKDEC : LREAL;
	LRJERKTIMEACC : LREAL;
	LRJERKTIMEDEC : LREAL;
END_VAR
VAR_OUTPUT
	DWSTATE : DWORD;
END_VAR
VAR_IN_OUT
	SCPROFILEDATA : L_MB1P_ProfileData;
	SCPROFILEPARAMETER : L_MB1P_ProfileParameter;
END_VAR
END_METHOD

METHOD CALCPROFILE_60B0_A0GTAMAX : BOOL
VAR_INPUT
	LRSTARTACC : LREAL;
	LRSTARTVEL : LREAL;
	LRMAXACC : LREAL;
	LRMAXDEC : LREAL;
	LRMAXVEL : LREAL;
	LRTARGETACC : LREAL;
	LRTARGETVEL : LREAL;
	LRTARGETPOS : LREAL;
	LRJERKACC : LREAL;
	LRJERKDEC : LREAL;
	LRJERKTIMEACC : LREAL;
	LRJERKTIMEDEC : LREAL;
END_VAR
VAR_IN_OUT
	SCPROFILEDATA : L_MB1P_ProfileData;
END_VAR
END_METHOD

METHOD CALCPROFILE_60B0_A0LTAMAX : BOOL
VAR_INPUT
	LRSTARTACC : LREAL;
	LRSTARTVEL : LREAL;
	LRMAXACC : LREAL;
	LRMAXDEC : LREAL;
	LRMAXVEL : LREAL;
	LRTARGETACC : LREAL;
	LRTARGETVEL : LREAL;
	LRTARGETPOS : LREAL;
	LRJERKACC : LREAL;
	LRJERKDEC : LREAL;
	LRJERKTIMEACC : LREAL;
	LRJERKTIMEDEC : LREAL;
END_VAR
VAR_IN_OUT
	SCPROFILEDATA : L_MB1P_ProfileData;
END_VAR
END_METHOD

METHOD CALCPROFILE_60C0 : BOOL
VAR_INPUT
	LRSTARTACC : LREAL;
	LRSTARTVEL : LREAL;
	LRMAXACC : LREAL;
	LRMAXDEC : LREAL;
	LRMAXVEL : LREAL;
	LRTARGETACC : LREAL;
	LRTARGETVEL : LREAL;
	LRTARGETPOS : LREAL;
	LRJERKACC : LREAL;
	LRJERKDEC : LREAL;
	LRJERKTIMEACC : LREAL;
	LRJERKTIMEDEC : LREAL;
END_VAR
VAR_OUTPUT
	DWSTATE : DWORD;
END_VAR
VAR_IN_OUT
	SCPROFILEDATA : L_MB1P_ProfileData;
	SCPROFILEPARAMETER : L_MB1P_ProfileParameter;
END_VAR
END_METHOD

METHOD CALCPROFILE_60D0 : BOOL
VAR_INPUT
	LRSTARTACC : LREAL;
	LRSTARTVEL : LREAL;
	LRMAXACC : LREAL;
	LRMAXDEC : LREAL;
	LRMAXVEL : LREAL;
	LRTARGETACC : LREAL;
	LRTARGETVEL : LREAL;
	LRTARGETPOS : LREAL;
	LRJERKACC : LREAL;
	LRJERKDEC : LREAL;
	LRJERKTIMEACC : LREAL;
	LRJERKTIMEDEC : LREAL;
END_VAR
VAR_OUTPUT
	DWSTATE : DWORD;
END_VAR
VAR_IN_OUT
	SCPROFILEDATA : L_MB1P_ProfileData;
	SCPROFILEPARAMETER : L_MB1P_ProfileParameter;
END_VAR
END_METHOD

METHOD CALCPROFILE_70A0 : BOOL
VAR_INPUT
	LRSTARTACC : LREAL;
	LRSTARTVEL : LREAL;
	LRMAXACC : LREAL;
	LRMAXDEC : LREAL;
	LRMAXVEL : LREAL;
	LRTARGETACC : LREAL;
	LRTARGETVEL : LREAL;
	LRTARGETPOS : LREAL;
	LRJERKACC : LREAL;
	LRJERKDEC : LREAL;
	LRJERKTIMEACC : LREAL;
	LRJERKTIMEDEC : LREAL;
	SCMAXPROFILEDATA : L_MB1P_IntProfileData;
	SCMINPROFILEDATA : L_MB1P_IntProfileData;
END_VAR
VAR_OUTPUT
	DWSTATE : DWORD;
END_VAR
VAR_IN_OUT
	SCPROFILEDATA : L_MB1P_ProfileData;
	SCPROFILEPARAMETER : L_MB1P_ProfileParameter;
END_VAR
END_METHOD

METHOD CALCPROFILE_70A0_SEARCHTIMEST5T7 : BOOL
VAR_INPUT
	LRSTARTACC : LREAL;
	LRSTARTVEL : LREAL;
	LRMAXACC : LREAL;
	LRMAXDEC : LREAL;
	LRMAXVEL : LREAL;
	LRTARGETACC : LREAL;
	LRTARGETVEL : LREAL;
	LRTARGETPOS : LREAL;
	LRJERKACC : LREAL;
	LRJERKDEC : LREAL;
	LRJERKTIMEACC : LREAL;
	LRJERKTIMEDEC : LREAL;
	T5_STARTVALUE : LREAL;
	T7_STARTVALUE : LREAL;
END_VAR
VAR_OUTPUT
	T5 : LREAL;
	T7 : LREAL;
END_VAR
END_METHOD

METHOD CALCPROFILE_70A0_A0LTAMAXT5T7 : BOOL
VAR_INPUT
	LRSTARTACC : LREAL;
	LRSTARTVEL : LREAL;
	LRMAXACC : LREAL;
	LRMAXDEC : LREAL;
	LRMAXVEL : LREAL;
	LRTARGETACC : LREAL;
	LRTARGETVEL : LREAL;
	LRTARGETPOS : LREAL;
	LRJERKACC : LREAL;
	LRJERKDEC : LREAL;
	LRJERKTIMEACC : LREAL;
	LRJERKTIMEDEC : LREAL;
	T5 : LREAL;
	T7 : LREAL;
END_VAR
VAR_OUTPUT
	A : ARRAY [1..4] OF LREAL;
END_VAR
VAR_IN_OUT
	SCPROFILEDATA : L_MB1P_ProfileData;
END_VAR
END_METHOD

METHOD CALCPROFILE_70B0 : BOOL
VAR_INPUT
	LRSTARTACC : LREAL;
	LRSTARTVEL : LREAL;
	LRMAXACC : LREAL;
	LRMAXDEC : LREAL;
	LRMAXVEL : LREAL;
	LRTARGETACC : LREAL;
	LRTARGETVEL : LREAL;
	LRTARGETPOS : LREAL;
	LRJERKACC : LREAL;
	LRJERKDEC : LREAL;
	LRJERKTIMEACC : LREAL;
	LRJERKTIMEDEC : LREAL;
	SCMAXPROFILEDATA : L_MB1P_IntProfileData;
	SCMINPROFILEDATA : L_MB1P_IntProfileData;
END_VAR
VAR_OUTPUT
	DWSTATE : DWORD;
END_VAR
VAR_IN_OUT
	SCPROFILEDATA : L_MB1P_ProfileData;
	SCPROFILEPARAMETER : L_MB1P_ProfileParameter;
END_VAR
END_METHOD

METHOD CALCPROFILE_70B0_SEARCHTIMEST5T7 : BOOL
VAR_INPUT
	LRSTARTACC : LREAL;
	LRSTARTVEL : LREAL;
	LRMAXACC : LREAL;
	LRMAXDEC : LREAL;
	LRMAXVEL : LREAL;
	LRTARGETACC : LREAL;
	LRTARGETVEL : LREAL;
	LRTARGETPOS : LREAL;
	LRJERKACC : LREAL;
	LRJERKDEC : LREAL;
	LRJERKTIMEACC : LREAL;
	LRJERKTIMEDEC : LREAL;
	T5_STARTVALUE : LREAL;
	T7_STARTVALUE : LREAL;
END_VAR
VAR_OUTPUT
	T5 : LREAL;
	T7 : LREAL;
END_VAR
END_METHOD

METHOD CALCPROFILE_70B0_A0LTAMAXT5T7 : BOOL
VAR_INPUT
	LRSTARTACC : LREAL;
	LRSTARTVEL : LREAL;
	LRMAXACC : LREAL;
	LRMAXDEC : LREAL;
	LRMAXVEL : LREAL;
	LRTARGETACC : LREAL;
	LRTARGETVEL : LREAL;
	LRTARGETPOS : LREAL;
	LRJERKACC : LREAL;
	LRJERKDEC : LREAL;
	LRJERKTIMEACC : LREAL;
	LRJERKTIMEDEC : LREAL;
	T5 : LREAL;
	T7 : LREAL;
END_VAR
VAR_OUTPUT
	A : ARRAY [1..4] OF LREAL;
END_VAR
VAR_IN_OUT
	SCPROFILEDATA : L_MB1P_ProfileData;
END_VAR
END_METHOD

METHOD CALCPROFILE_80A0 : BOOL
VAR_INPUT
	LRSTARTACC : LREAL;
	LRSTARTVEL : LREAL;
	LRMAXACC : LREAL;
	LRMAXDEC : LREAL;
	LRMAXVEL : LREAL;
	LRTARGETACC : LREAL;
	LRTARGETVEL : LREAL;
	LRTARGETPOS : LREAL;
	LRJERKACC : LREAL;
	LRJERKDEC : LREAL;
	LRJERKTIMEACC : LREAL;
	LRJERKTIMEDEC : LREAL;
	SCMAXPROFILEDATA : L_MB1P_IntProfileData;
	SCMINPROFILEDATA : L_MB1P_IntProfileData;
END_VAR
VAR_OUTPUT
	DWSTATE : DWORD;
END_VAR
VAR_IN_OUT
	SCPROFILEDATA : L_MB1P_ProfileData;
	SCPROFILEPARAMETER : L_MB1P_ProfileParameter;
END_VAR
END_METHOD

METHOD CALCPROFILE_80A0_A0GTAMAXT5T7 : BOOL
VAR_INPUT
	LRSTARTACC : LREAL;
	LRSTARTVEL : LREAL;
	LRMAXACC : LREAL;
	LRMAXDEC : LREAL;
	LRMAXVEL : LREAL;
	LRTARGETACC : LREAL;
	LRTARGETVEL : LREAL;
	LRTARGETPOS : LREAL;
	LRJERKACC : LREAL;
	LRJERKDEC : LREAL;
	LRJERKTIMEACC : LREAL;
	LRJERKTIMEDEC : LREAL;
	T5 : LREAL;
	T7 : LREAL;
END_VAR
VAR_IN_OUT
	SCPROFILEDATA : L_MB1P_ProfileData;
END_VAR
END_METHOD

METHOD CALCPROFILE_80A0_A0GTAMAX_SEARCHTIMEST5T7 : BOOL
VAR_INPUT
	LRSTARTACC : LREAL;
	LRSTARTVEL : LREAL;
	LRMAXACC : LREAL;
	LRMAXDEC : LREAL;
	LRMAXVEL : LREAL;
	LRTARGETACC : LREAL;
	LRTARGETVEL : LREAL;
	LRTARGETPOS : LREAL;
	LRJERKACC : LREAL;
	LRJERKDEC : LREAL;
	LRJERKTIMEACC : LREAL;
	LRJERKTIMEDEC : LREAL;
	T5_STARTVALUE : LREAL;
	T7_STARTVALUE : LREAL;
END_VAR
VAR_OUTPUT
	T5 : LREAL;
	T7 : LREAL;
END_VAR
END_METHOD

METHOD CALCPROFILE_80A0_A0LTAMAXT5T7 : BOOL
VAR_INPUT
	LRSTARTACC : LREAL;
	LRSTARTVEL : LREAL;
	LRMAXACC : LREAL;
	LRMAXDEC : LREAL;
	LRMAXVEL : LREAL;
	LRTARGETACC : LREAL;
	LRTARGETVEL : LREAL;
	LRTARGETPOS : LREAL;
	LRJERKACC : LREAL;
	LRJERKDEC : LREAL;
	LRJERKTIMEACC : LREAL;
	LRJERKTIMEDEC : LREAL;
	T5 : LREAL;
	T7 : LREAL;
END_VAR
VAR_IN_OUT
	SCPROFILEDATA : L_MB1P_ProfileData;
END_VAR
END_METHOD

METHOD CALCPROFILE_80A0_A0LTAMAX_SEARCHTIMEST5T7 : BOOL
VAR_INPUT
	LRSTARTACC : LREAL;
	LRSTARTVEL : LREAL;
	LRMAXACC : LREAL;
	LRMAXDEC : LREAL;
	LRMAXVEL : LREAL;
	LRTARGETACC : LREAL;
	LRTARGETVEL : LREAL;
	LRTARGETPOS : LREAL;
	LRJERKACC : LREAL;
	LRJERKDEC : LREAL;
	LRJERKTIMEACC : LREAL;
	LRJERKTIMEDEC : LREAL;
	T5_STARTVALUE : LREAL;
	T7_STARTVALUE : LREAL;
END_VAR
VAR_OUTPUT
	T5 : LREAL;
	T7 : LREAL;
END_VAR
END_METHOD

METHOD CALCPROFILE_80B0 : BOOL
VAR_INPUT
	LRSTARTACC : LREAL;
	LRSTARTVEL : LREAL;
	LRMAXACC : LREAL;
	LRMAXDEC : LREAL;
	LRMAXVEL : LREAL;
	LRTARGETACC : LREAL;
	LRTARGETVEL : LREAL;
	LRTARGETPOS : LREAL;
	LRJERKACC : LREAL;
	LRJERKDEC : LREAL;
	LRJERKTIMEACC : LREAL;
	LRJERKTIMEDEC : LREAL;
	SCMAXPROFILEDATA : L_MB1P_IntProfileData;
	SCMINPROFILEDATA : L_MB1P_IntProfileData;
END_VAR
VAR_OUTPUT
	DWSTATE : DWORD;
END_VAR
VAR_IN_OUT
	SCPROFILEDATA : L_MB1P_ProfileData;
	SCPROFILEPARAMETER : L_MB1P_ProfileParameter;
END_VAR
END_METHOD

METHOD CALCPROFILE_80B0_A0GTAMAX_SEARCHTIMEST5T7 : BOOL
VAR_INPUT
	LRSTARTACC : LREAL;
	LRSTARTVEL : LREAL;
	LRMAXACC : LREAL;
	LRMAXDEC : LREAL;
	LRMAXVEL : LREAL;
	LRTARGETACC : LREAL;
	LRTARGETVEL : LREAL;
	LRTARGETPOS : LREAL;
	LRJERKACC : LREAL;
	LRJERKDEC : LREAL;
	LRJERKTIMEACC : LREAL;
	LRJERKTIMEDEC : LREAL;
	T5_STARTVALUE : LREAL;
	T7_STARTVALUE : LREAL;
END_VAR
VAR_OUTPUT
	T5 : LREAL;
	T7 : LREAL;
END_VAR
END_METHOD

METHOD CALCPROFILE_80B0_A0GTAMAXT5T7 : BOOL
VAR_INPUT
	LRSTARTACC : LREAL;
	LRSTARTVEL : LREAL;
	LRMAXACC : LREAL;
	LRMAXDEC : LREAL;
	LRMAXVEL : LREAL;
	LRTARGETACC : LREAL;
	LRTARGETVEL : LREAL;
	LRTARGETPOS : LREAL;
	LRJERKACC : LREAL;
	LRJERKDEC : LREAL;
	LRJERKTIMEACC : LREAL;
	LRJERKTIMEDEC : LREAL;
	T5 : LREAL;
	T7 : LREAL;
END_VAR
VAR_IN_OUT
	SCPROFILEDATA : L_MB1P_ProfileData;
END_VAR
END_METHOD

METHOD CALCPROFILE_80B0_A0LTAMAXT5T7 : BOOL
VAR_INPUT
	LRSTARTACC : LREAL;
	LRSTARTVEL : LREAL;
	LRMAXACC : LREAL;
	LRMAXDEC : LREAL;
	LRMAXVEL : LREAL;
	LRTARGETACC : LREAL;
	LRTARGETVEL : LREAL;
	LRTARGETPOS : LREAL;
	LRJERKACC : LREAL;
	LRJERKDEC : LREAL;
	LRJERKTIMEACC : LREAL;
	LRJERKTIMEDEC : LREAL;
	T5 : LREAL;
	T7 : LREAL;
END_VAR
VAR_IN_OUT
	SCPROFILEDATA : L_MB1P_ProfileData;
END_VAR
END_METHOD

METHOD CALCPROFILE_80B0_A0LTAMAX_SEARCHTIMEST5T7 : BOOL
VAR_INPUT
	LRSTARTACC : LREAL;
	LRSTARTVEL : LREAL;
	LRMAXACC : LREAL;
	LRMAXDEC : LREAL;
	LRMAXVEL : LREAL;
	LRTARGETACC : LREAL;
	LRTARGETVEL : LREAL;
	LRTARGETPOS : LREAL;
	LRJERKACC : LREAL;
	LRJERKDEC : LREAL;
	LRJERKTIMEACC : LREAL;
	LRJERKTIMEDEC : LREAL;
	T5_STARTVALUE : LREAL;
	T7_STARTVALUE : LREAL;
END_VAR
VAR_OUTPUT
	T5 : LREAL;
	T7 : LREAL;
END_VAR
END_METHOD

METHOD CALCPROFILE_80C0 : BOOL
VAR_INPUT
	LRSTARTACC : LREAL;
	LRSTARTVEL : LREAL;
	LRMAXACC : LREAL;
	LRMAXDEC : LREAL;
	LRMAXVEL : LREAL;
	LRTARGETACC : LREAL;
	LRTARGETVEL : LREAL;
	LRTARGETPOS : LREAL;
	LRJERKACC : LREAL;
	LRJERKDEC : LREAL;
	LRJERKTIMEACC : LREAL;
	LRJERKTIMEDEC : LREAL;
	SCMAXPROFILEDATA : L_MB1P_IntProfileData;
	SCMINPROFILEDATA : L_MB1P_IntProfileData;
END_VAR
VAR_OUTPUT
	DWSTATE : DWORD;
END_VAR
VAR_IN_OUT
	SCPROFILEDATA : L_MB1P_ProfileData;
	SCPROFILEPARAMETER : L_MB1P_ProfileParameter;
END_VAR
END_METHOD

METHOD CALCPROFILE_80C0_SEARCHTIMEST5T7 : BOOL
VAR_INPUT
	LRSTARTACC : LREAL;
	LRSTARTVEL : LREAL;
	LRMAXACC : LREAL;
	LRMAXDEC : LREAL;
	LRMAXVEL : LREAL;
	LRTARGETACC : LREAL;
	LRTARGETVEL : LREAL;
	LRTARGETPOS : LREAL;
	LRJERKACC : LREAL;
	LRJERKDEC : LREAL;
	LRJERKTIMEACC : LREAL;
	LRJERKTIMEDEC : LREAL;
	T5_STARTVALUE : LREAL;
	T7_STARTVALUE : LREAL;
END_VAR
VAR_OUTPUT
	T5 : LREAL;
	T7 : LREAL;
END_VAR
END_METHOD

METHOD CALCPROFILE_80C0_A0LTAMAXT5T7 : BOOL
VAR_INPUT
	LRSTARTACC : LREAL;
	LRSTARTVEL : LREAL;
	LRMAXACC : LREAL;
	LRMAXDEC : LREAL;
	LRMAXVEL : LREAL;
	LRTARGETACC : LREAL;
	LRTARGETVEL : LREAL;
	LRTARGETPOS : LREAL;
	LRJERKACC : LREAL;
	LRJERKDEC : LREAL;
	LRJERKTIMEACC : LREAL;
	LRJERKTIMEDEC : LREAL;
	T5 : LREAL;
	T7 : LREAL;
END_VAR
VAR_IN_OUT
	SCPROFILEDATA : L_MB1P_ProfileData;
END_VAR
END_METHOD

METHOD CALCPROFILE_80D0 : BOOL
VAR_INPUT
	LRSTARTACC : LREAL;
	LRSTARTVEL : LREAL;
	LRMAXACC : LREAL;
	LRMAXDEC : LREAL;
	LRMAXVEL : LREAL;
	LRTARGETACC : LREAL;
	LRTARGETVEL : LREAL;
	LRTARGETPOS : LREAL;
	LRJERKACC : LREAL;
	LRJERKDEC : LREAL;
	LRJERKTIMEACC : LREAL;
	LRJERKTIMEDEC : LREAL;
	SCMAXPROFILEDATA : L_MB1P_IntProfileData;
	SCMINPROFILEDATA : L_MB1P_IntProfileData;
END_VAR
VAR_OUTPUT
	DWSTATE : DWORD;
END_VAR
VAR_IN_OUT
	SCPROFILEDATA : L_MB1P_ProfileData;
	SCPROFILEPARAMETER : L_MB1P_ProfileParameter;
END_VAR
END_METHOD

METHOD CALCPROFILE_80D0_SEARCHTIMEST5T7 : BOOL
VAR_INPUT
	LRSTARTACC : LREAL;
	LRSTARTVEL : LREAL;
	LRMAXACC : LREAL;
	LRMAXDEC : LREAL;
	LRMAXVEL : LREAL;
	LRTARGETACC : LREAL;
	LRTARGETVEL : LREAL;
	LRTARGETPOS : LREAL;
	LRJERKACC : LREAL;
	LRJERKDEC : LREAL;
	LRJERKTIMEACC : LREAL;
	LRJERKTIMEDEC : LREAL;
	T5_STARTVALUE : LREAL;
	T7_STARTVALUE : LREAL;
END_VAR
VAR_OUTPUT
	T5 : LREAL;
	T7 : LREAL;
END_VAR
END_METHOD

METHOD CALCPROFILE_80D0_A0LTAMAXT5T7 : BOOL
VAR_INPUT
	LRSTARTACC : LREAL;
	LRSTARTVEL : LREAL;
	LRMAXACC : LREAL;
	LRMAXDEC : LREAL;
	LRMAXVEL : LREAL;
	LRTARGETACC : LREAL;
	LRTARGETVEL : LREAL;
	LRTARGETPOS : LREAL;
	LRJERKACC : LREAL;
	LRJERKDEC : LREAL;
	LRJERKTIMEACC : LREAL;
	LRJERKTIMEDEC : LREAL;
	T5 : LREAL;
	T7 : LREAL;
END_VAR
VAR_IN_OUT
	SCPROFILEDATA : L_MB1P_ProfileData;
END_VAR
END_METHOD

METHOD CALCPROFILE_80E0 : BOOL
VAR_INPUT
	LRSTARTACC : LREAL;
	LRSTARTVEL : LREAL;
	LRMAXACC : LREAL;
	LRMAXDEC : LREAL;
	LRMAXVEL : LREAL;
	LRTARGETACC : LREAL;
	LRTARGETVEL : LREAL;
	LRTARGETPOS : LREAL;
	LRJERKACC : LREAL;
	LRJERKDEC : LREAL;
	LRJERKTIMEACC : LREAL;
	LRJERKTIMEDEC : LREAL;
	SCMAXPROFILEDATA : L_MB1P_IntProfileData;
	SCMINPROFILEDATA : L_MB1P_IntProfileData;
END_VAR
VAR_OUTPUT
	DWSTATE : DWORD;
END_VAR
VAR_IN_OUT
	SCPROFILEDATA : L_MB1P_ProfileData;
	SCPROFILEPARAMETER : L_MB1P_ProfileParameter;
END_VAR
END_METHOD

METHOD CALCPROFILE_80E0_PROFILEDATA : BOOL
VAR_INPUT
	LRSTARTACC : LREAL;
	LRSTARTVEL : LREAL;
	LRMAXACC : LREAL;
	LRMAXDEC : LREAL;
	LRMAXVEL : LREAL;
	LRTARGETACC : LREAL;
	LRTARGETVEL : LREAL;
	LRTARGETPOS : LREAL;
	LRJERKACC : LREAL;
	LRJERKDEC : LREAL;
	LRJERKTIMEACC : LREAL;
	LRJERKTIMEDEC : LREAL;
	T5 : LREAL;
	T7 : LREAL;
END_VAR
VAR_IN_OUT
	SCPROFILEDATA : L_MB1P_ProfileData;
END_VAR
END_METHOD

METHOD CALCPROFILE_80E0_SEARCHTIMEST5T7 : BOOL
VAR_INPUT
	LRSTARTACC : LREAL;
	LRSTARTVEL : LREAL;
	LRMAXACC : LREAL;
	LRMAXDEC : LREAL;
	LRMAXVEL : LREAL;
	LRTARGETACC : LREAL;
	LRTARGETVEL : LREAL;
	LRTARGETPOS : LREAL;
	LRJERKACC : LREAL;
	LRJERKDEC : LREAL;
	LRJERKTIMEACC : LREAL;
	LRJERKTIMEDEC : LREAL;
	T5_STARTVALUE : LREAL;
	T7_STARTVALUE : LREAL;
END_VAR
VAR_OUTPUT
	T5 : LREAL;
	T7 : LREAL;
END_VAR
END_METHOD

METHOD CALCPROFILE_80F0 : BOOL
VAR_INPUT
	LRSTARTACC : LREAL;
	LRSTARTVEL : LREAL;
	LRMAXACC : LREAL;
	LRMAXDEC : LREAL;
	LRMAXVEL : LREAL;
	LRTARGETACC : LREAL;
	LRTARGETVEL : LREAL;
	LRTARGETPOS : LREAL;
	LRJERKACC : LREAL;
	LRJERKDEC : LREAL;
	LRJERKTIMEACC : LREAL;
	LRJERKTIMEDEC : LREAL;
	SCMAXPROFILEDATA : L_MB1P_IntProfileData;
	SCMINPROFILEDATA : L_MB1P_IntProfileData;
END_VAR
VAR_OUTPUT
	DWSTATE : DWORD;
END_VAR
VAR_IN_OUT
	SCPROFILEDATA : L_MB1P_ProfileData;
	SCPROFILEPARAMETER : L_MB1P_ProfileParameter;
END_VAR
END_METHOD

METHOD CALCPROFILE_80F0_PROFILEDATA : BOOL
VAR_INPUT
	LRSTARTACC : LREAL;
	LRSTARTVEL : LREAL;
	LRMAXACC : LREAL;
	LRMAXDEC : LREAL;
	LRMAXVEL : LREAL;
	LRTARGETACC : LREAL;
	LRTARGETVEL : LREAL;
	LRTARGETPOS : LREAL;
	LRJERKACC : LREAL;
	LRJERKDEC : LREAL;
	LRJERKTIMEACC : LREAL;
	LRJERKTIMEDEC : LREAL;
	T5 : LREAL;
	T7 : LREAL;
END_VAR
VAR_IN_OUT
	SCPROFILEDATA : L_MB1P_ProfileData;
END_VAR
END_METHOD

METHOD CALCPROFILE_80F0_SEARCHTIMEST5T7 : BOOL
VAR_INPUT
	LRSTARTACC : LREAL;
	LRSTARTVEL : LREAL;
	LRMAXACC : LREAL;
	LRMAXDEC : LREAL;
	LRMAXVEL : LREAL;
	LRTARGETACC : LREAL;
	LRTARGETVEL : LREAL;
	LRTARGETPOS : LREAL;
	LRJERKACC : LREAL;
	LRJERKDEC : LREAL;
	LRJERKTIMEACC : LREAL;
	LRJERKTIMEDEC : LREAL;
	T5_STARTVALUE : LREAL;
	T7_STARTVALUE : LREAL;
END_VAR
VAR_OUTPUT
	T5 : LREAL;
	T7 : LREAL;
END_VAR
END_METHOD

(* ---- L_MB1P_POSPROFILERCLUTCH.fb ---- *)
FUNCTION_BLOCK L_MB1P_POSPROFILERCLUTCH
VAR_INPUT
	XENABLE : BOOL;
	XSYNCPOS : BOOL;
	XEXECUTEGAP : BOOL;
	XAUXEXECUTEGAP : BOOL;
	LRTASKCYCLETIME : LREAL := 0.001;
	LRSLAVESYNCOUTPOS : LREAL;
	LRCYCMASTERPOS : LREAL;
	LRCYCMASTERVEL : LREAL;
	LRCYCMASTERACC : LREAL;
	LRSETSLAVEPOS : LREAL;
	LRSETSLAVEVEL : LREAL;
	LRSETSLAVEACC : LREAL;
	LRJERK : LREAL := 10000;
	LRMAXACC : LREAL := 100;
	LRMAXDEC : LREAL := 100;
	LRMAXVEL : LREAL := 10;
END_VAR
VAR_OUTPUT
	XBUSY : BOOL;
	XDONE : BOOL;
	XACCDECSYNC : BOOL;
	XPOSSYNCHRONISED : BOOL;
	XERROR : BOOL;
	EERRORID : WORD;
	LRSETSLAVEPOSOUT : LREAL;
	LRSETSLAVEVELOUT : LREAL;
	LRSETSLAVEACCOUT : LREAL;
END_VAR
VAR
	FB_POSPROFILERPOS : L_MC1P_PosProfiler;
	SCPROFILEPARAMETER : L_MC1P_ProfileParameter;
	WSTEPPER : WORD;
	XEXECUTEPOSPROFILER : BOOL;
	LRSLAVESYNCOUTPOS_INT : LREAL;
	XAUXEXECUTEPROFILE : BOOL;
	XEXECUTEPROFILE : BOOL;
	LRSETPOSPROFILER : LREAL;
	LRSETACCPROFILER : LREAL;
	LRSETVELPROFILER : LREAL;
	LRCYCMASTERPOS_INT : LREAL;
	LRCYCMASTERVEL_INT : LREAL;
	LRCYCMASTERACC_INT : LREAL;
	XPOSSYNCHRONISED_INT : BOOL;
	XEXECUTEGAPOLD : BOOL;
	XAUXEXECUTEGAPOLD : BOOL;
	XENABLEOLD : BOOL;
	LRCYCMASTERPOS_OLD : LREAL;
	LRTOLERANCE : LREAL;
END_VAR
END_FUNCTION_BLOCK

METHOD CALL_ERRORHANDLER
END_METHOD

METHOD CALL_FBMETHODES
END_METHOD

METHOD CALL_FB_POSPROFILERPOS
END_METHOD

METHOD CALL_FB_POSPROFILERPOSINPUTS
END_METHOD

METHOD CALL_OUTPUTS
END_METHOD

METHOD CALL_PROFILEPARAMETER
END_METHOD

METHOD CALL_RESETCOMMANDS
END_METHOD

METHOD CALL_RESETOUTPUTS
END_METHOD

METHOD CALL_STATEMACHINE
END_METHOD

(* ---- L_MB1P_POSPROFILERCLUTCHSTATE.fb ---- *)
FUNCTION_BLOCK L_MB1P_POSPROFILERCLUTCHSTATE EXTENDS L_MB1P_PosProfilerClutch
VAR_INPUT
	XSYNCOUTINSTANT : BOOL;
	XMOVETOTARGETPOS : BOOL;
	LRTARGETPOS : LREAL;
	EDIRECTION : L_MC2P_ClutchDirection := L_MC2P_ClutchDirection.mcCurrentDirection;
	LRAXESCYCLELENGTH : LREAL := 360;
	EAXESTRAVERSINGRANGE : L_MC1P_TraversingRange;
	LRPOSITIONINGJERK : LREAL;
	LRPOSITIONINGACC : LREAL;
	LRPOSITIONINGDEC : LREAL;
	LRPOSITIONINGVEL : LREAL;
	LRSYNCOUTINSTANTJERK : LREAL;
	LRSYNCOUTINSTANTDEC : LREAL;
	ROVERRIDEVEL : REAL := 1.0;
	ROVERRIDEACC : REAL := 1.0;
	ROVERRIDEDEC : REAL := 1.0;
END_VAR
VAR_OUTPUT
	XREVERSING : BOOL;
	XPOSITIONING : BOOL;
	XINPOSITION : BOOL;
END_VAR
VAR
	XREVERSING_INT : BOOL;
	WMODE : WORD;
	XSYNCOUTINSTANT_OLD : BOOL;
	XMOVETOTARGETPOS_OLD : BOOL;
	XPOSMODE_INT : BOOL;
	LRTASKCYCLETIME_INT : LREAL;
	LRAXESCYCLELENGTH_INT : LREAL;
	LRTARGETPOS_INT : LREAL;
	LRTARGETPOS_LOCK : LREAL;
	LRTOLERANCEVEL : LREAL;
	LRTOLERANCEACC : LREAL;
	LRACCDIST : LREAL;
	XVELTRACE : BOOL;
	WVELTRACESTEPPER : WORD;
	LRSETACC_PROFILERPOS : LREAL;
	LRPOSPROFILERSPEED_ABS : LREAL;
	WREVERSINGVELMODE : WORD;
	LRVELZERROTOLERANZ : LREAL;
	LRSETSLAVEVELOUT_OLD : LREAL;
END_VAR
END_FUNCTION_BLOCK

METHOD CALL_CALCTARGETPOS
VAR_INPUT
	LRTARGETPOS : LREAL;
END_VAR
END_METHOD

METHOD CALL_CALCTOLERANCE
END_METHOD

METHOD CALL_CALCLRCYCMASTERPOS
END_METHOD

METHOD CALL_ERRORHANDLER
END_METHOD

METHOD CALL_FBMETHODES
END_METHOD

METHOD CALL_FB_POSPROFILERPOS
END_METHOD

METHOD CALL_FB_POSPROFILERPOSINPUTS
END_METHOD

METHOD CALL_OUTPUTS
END_METHOD

METHOD CALL_PROFILEPARAMETER
END_METHOD

METHOD CALL_PROFILEPARAMETERACCDECINMODE2
END_METHOD

METHOD CALL_RESETCOMMANDS
END_METHOD

METHOD CALL_RESETOUTPUTS
END_METHOD

METHOD CALL_STATEMACHINE
END_METHOD

(* ---- L_MB1P_PREPARATIONPATH_LM.fb ---- *)
FUNCTION_BLOCK L_MB1P_PREPARATIONPATH_LM
VAR_INPUT
	XEXECUTE : BOOL;
	XSINGLESTEP : BOOL;
	ALRSTARTPOSITION : ARRAY [1..12] OF LREAL;
	LRSTARTBLENDINGRADIUS : LREAL;
	XSTARTHALT : BOOL;
	LRPATHJERK : LREAL;
	XECOCPUMODE : BOOL;
END_VAR
VAR_OUTPUT
	XERROR : BOOL;
	EERRORID : L_IE1P_Error;
	XBUSY : BOOL;
	XDONE : BOOL;
	BYNUMOFPOINTS : BYTE;
	BYNUMOFHALT : BYTE;
	AXHALT : ARRAY [0..10] OF BOOL;
	ALRPROFILEPOINTS : ARRAY [1..10] OF ARRAY [1..12] OF LREAL;
	EENDCOORDSYSTEM : L_MC4P_CoordSystem := L_MC4P_CoordSystem.MCS;
	ALRENDPOSITION : ARRAY [1..12] OF LREAL;
	LRENDBLENDINGRADIUS : LREAL;
	XENDHALT : BOOL;
END_VAR
VAR_IN_OUT
	AXESGROUP : AXES_GROUP_KIN;
	ASCPROFILEPAR : ARRAY [1..10] OF L_TT1P_scProfilePar;
	MC_MOVELINABS : ARRAY [1..10] OF MC_MoveLinearAbsolute;
END_VAR
VAR
	WSTATE : WORD := 0;
	AXCALCPATHLEGTHBETWEENPOINTS : ARRAY [1..11] OF BOOL;
	ALRPATHLEGTHBETWEENPOINTS : ARRAY [1..11] OF LREAL;
	XSINGLESTEP_INT : BOOL;
	LRBLENDINGRADIUS_INT : LREAL;
	BYNUMOFPOINTS_LOCK : BYTE;
	XCALCINTERMEDIANTEPOINT : BOOL;
	XCPUECOMODEEXECUTE : BOOL;
	IPOINTNO : INT;
	IFORCNT : INT;
	IFORCNT2 : INT;
	LRTMP : LREAL;
	LRTMP1 : LREAL;
	LRTMP2 : LREAL;
	XERRORINVALIDPROFILE : BOOL;
	XERROR_INVALIDCOORDSYSTEM : BOOL;
	XERROR_INTERNAL : BOOL;
	XEXECUTE_OLD : BOOL;
	C_BYMAXTARGETPOINTS : BYTE := 10;
END_VAR
END_FUNCTION_BLOCK

METHOD CALL_ERRORHANDLER
END_METHOD

METHOD CALL_FBMETHODS
END_METHOD

METHOD CALL_OUTPUT
END_METHOD

METHOD CALL_RESETCOMMANDS
END_METHOD

METHOD CALL_RESETFB
END_METHOD

METHOD CALL_RESETOUTPUT
END_METHOD

METHOD CALL_STATEMACHINE
END_METHOD

METHOD GET_LRTARTGETPOSITION : LREAL
VAR_INPUT
	IAXISID : INT;
	IPOINTNO : INT;
END_VAR
END_METHOD

METHOD CALL_INIT
END_METHOD

(* ---- L_MB1P_SIMPLEPOSABORTCORRECTION.fb ---- *)
FUNCTION_BLOCK L_MB1P_SIMPLEPOSABORTCORRECTION
VAR_INPUT
	XENABLE : BOOL;
	LRCYCLETIME : LREAL;
	XABORTFROMPOSCTRL : BOOL;
	LRMAXACC : LREAL;
	LRACTVELFROMPOSCTRL : LREAL;
	LRSIMPLEPOSUNLIMITED : LREAL;
END_VAR
VAR_OUTPUT
	XABORTPROFILEFINISHED : BOOL;
	LRPOSOUT : LREAL;
END_VAR
VAR
	T_NORM_FAK : LREAL;
	T_NORM : LREAL;
	T_REAL : LREAL;
	LRSTARTPOS : LREAL;
	LRSTARTVEL : LREAL;
	R_EDGE_ABORTFROMPOSCTRL : R_TRIG;
	F_EDGE_ABORTFROMPOSCTRL : F_TRIG;
END_VAR
END_FUNCTION_BLOCK

(* ---- L_MB1P_SIMPLEPOSBASE.fb ---- *)
FUNCTION_BLOCK L_MB1P_SIMPLEPOSBASE
VAR_INPUT
	XENABLE : BOOL;
	XEXECUTE : BOOL;
	XABORTPROFILE : BOOL;
	LRCORRECTION : LREAL;
	LRMAXVELPOS : LREAL := 10;
	LRMAXVELNEG : LREAL := 10;
	LRACCDEC : LREAL := 100;
	EPROFILETYPE : L_MB1P_ProfileType := 0;
END_VAR
VAR_OUTPUT
	LRPOSOUTUNLIMITED : LREAL;
	LRRESIDUALOFFSET : LREAL;
	LRSPEEDOUT : LREAL;
	XPROFILEFAILED : BOOL;
	XPROFILEABORTED : BOOL;
	XINTARGET : BOOL;
	XBUSY : BOOL;
	DISTATE : DINT;
END_VAR
VAR_IN_OUT
	AXIS : Axis_REF;
END_VAR
VAR
	L_SDINTEGRATE1 : L_USPP_Integrate;
	R_TRIG1 : R_TRIG;
	R_TRIG2 : R_TRIG;
	F_TRIG2 : F_TRIG;
	F_TRIG3 : F_TRIG;
	DWPOSMODE : DWORD := 1;
	DWDISABLEMODE : DWORD;
	LRRAMPDISTANCE : LREAL;
	LRDELTAY : LREAL;
	LRBASICPOSITION : LREAL;
	BYSTEP : BYTE;
	BNEGSPEEDSELECTED : BOOL;
	LRXNORM : LREAL;
	LRPOSOUTOLD : LREAL;
	N : INT;
	LRMAXSPEEDINTERN : LREAL;
	LRMAXSPEEDNEG : LREAL;
	LRMAXSPEEDPOS : LREAL;
	LRSTARTPOSITION : LREAL;
	XSAVESTARTPOSITION : BOOL;
	LRPOSOUT : LREAL;
	LRPOSOUTOLDTEST : LREAL;
	LRPOSTEST : LREAL;
	XENDOFPROFILE : BOOL;
END_VAR
END_FUNCTION_BLOCK

METHOD A01_PROFILECONTROL
END_METHOD

METHOD A02_POLYNOMIAL4THORDER
END_METHOD

METHOD A03_POLYNOMIAL2NDORDER
END_METHOD

METHOD A04_POLYNOMIAL5THORDER
END_METHOD

(* ---- L_MB1P_SIMPLEPOSSETOFFSET.fb ---- *)
FUNCTION_BLOCK L_MB1P_SIMPLEPOSSETOFFSET
VAR_INPUT
	XENABLE : BOOL;
	LRCYCMASTERPOS : LREAL;
	LRCYCMASTERVEL : LREAL;
	LRCYCMASTERACC : LREAL;
	LRSETOFFSET : LREAL;
	XLOADOFFSET : BOOL;
	DWNUMERATOR : DWORD := 1;
	DWDENOMINATOR : DWORD := 1;
	EDIRECTION : L_TF1P_Direction;
	EPROFILETYPE : L_MB1P_ProfileType := 0;
	LRVELPOS : LREAL := 100.0;
	LRVELNEG : LREAL := 100.0;
	LRACCDEC : LREAL := 1000.0;
END_VAR
VAR_OUTPUT
	XBUSY : BOOL;
	XDONE : BOOL;
	XERROR : BOOL;
	EERRORID : WORD;
	LROFFSET : LREAL;
	LRSETOFFSETVELOUT : LREAL;
END_VAR
VAR_IN_OUT
	MASTERAXIS : AXIS_REF;
	SLAVEAXIS : AXIS_REF;
END_VAR
VAR
	WSTATEMASHINESIMPLEPOS : WORD := 0;
	LRSMDELTAPOS : LREAL;
	LRSIMPLEPOSOFFSET : LREAL;
	LRSALVEVELBAND : LREAL;
	LRABORTSTARTVEL : LREAL;
	LRSMSETOFFSET_OLD : LREAL;
	LRFACTOR : LREAL;
	LRLOADRESTOFFSET_INT : LREAL;
	LRVELPOS_INT : LREAL := 100.0;
	LRVELNEG_INT : LREAL := 100.0;
	LRACCDEC_INT : LREAL := 1000.0;
	XERRORINVALIDVELPOS : BOOL;
	XERRORINVALIDVELNEG : BOOL;
	XERRORINVALIDACCDEC : BOOL;
	XENABLE_OLD : BOOL;
	LROFFSET_OLD : LREAL;
	SIMPLEPOSITIONING : L_MB1P_SimplePosBase;
	ABORTPOSCTRLCORRECT : L_MB1P_SimplePosAbortCorrection;
END_VAR
END_FUNCTION_BLOCK

METHOD CALL_CALCFACTOR
END_METHOD

METHOD CALL_ERRORHANDLER
END_METHOD

METHOD CALL_FBMETHODS
END_METHOD

METHOD CALL_OUTPUT
END_METHOD

METHOD CALL_RESETCOMMANDS
END_METHOD

METHOD CALL_RESETOUTPUT
END_METHOD

METHOD CALL_SIMPLEPOS
END_METHOD

METHOD CALL_SIMPLEPOS_ABORTPOSCTRLCORRECT
END_METHOD

METHOD CALL_SIMPLEPOS_OFFSET
END_METHOD

METHOD CALL_STATEMASHINE
END_METHOD

(* ---- L_MB1P_STACK.fb ---- *)
FUNCTION_BLOCK L_MB1P_STACK
VAR_INPUT
	XENABLE : BOOL;
	XLOADTPPOS : BOOL;
	XLOADCYCSETPOS : BOOL;
	XTAKEPOS : BOOL;
	LRTPPOS : LREAL;
	LRCYCSETPOS : LREAL;
	LRCYCSETVEL : LREAL;
	LRPERIOD : LREAL;
	LRMINTPDIST : LREAL;
END_VAR
VAR_OUTPUT
	XBUSY : BOOL;
	XSTACKISFULL : BOOL;
	XSTACKISEMPTY : BOOL;
	LRPOSOUT : LREAL;
	LRDISTOUT : LREAL;
	LRSETDISTOUT : LREAL;
	XPOSPERIODOVERRUNPOS : BOOL;
	XPOSPERIODOVERRUNNEG : BOOL;
	UISTACKSTARTPOS : UINT := 0;
	UISTACKFILLSTATE : UINT := 0;
	ALRSTACKSAVEPOS : ARRAY [1..gc_uiStackLength] OF LREAL;
	AUIPERIODCNTRPOS : ARRAY [1..gc_uiStackLength] OF UINT;
	UIPERIODCNTR : UINT;
	LRTPDIST : LREAL;
	XPOSRECEIVED : BOOL;
	XPOSOUTOFWINDOW : BOOL;
	XWINDOWOPEN : BOOL;
END_VAR
VAR
	XSTACKVALUEVALID : BOOL;
	LRLATESTSAVEPOS : LREAL;
	UILATESTPERIODCNTRPOS : UINT;
	UICTR : UINT := 0;
	UIVARTEMP : UINT;
	XENABLE_OLD : BOOL;
	XLOADTPPOS_OLD : BOOL;
	XLOADCYCSETPOS_OLD : BOOL;
	XTAKEPOS_OLD : BOOL;
	XFIRSTLOADPOS : BOOL;
	LRCYCSETPOS_SAVE : LREAL;
	LRSETPOSDIFF : LREAL;
	XTAKEPOS_ACTIVE : BOOL;
	LRTEMPDIST : LREAL;
	LRCYCSETPOS_OLD : LREAL;
	FB_CHECKMODULOOVERRUN : L_MB1P_CheckModuloOverrun;
	GC_UISTACKLENGTH : UINT := 100;
END_VAR
END_FUNCTION_BLOCK

METHOD CALL_CNTRMODULOOVERRUN
VAR_IN_OUT
	LRCYCSETPOS : LREAL;
END_VAR
END_METHOD

METHOD CALL_FB_CHECKMODULOOVERRUN
VAR_IN_OUT
	LRCYCSETPOS : LREAL;
	LRCYCSETVEL : LREAL;
END_VAR
END_METHOD

METHOD CALL_RESETCOMMANDS
END_METHOD

METHOD CALL_RESETOUTPUT
END_METHOD

METHOD CALL_STACK
END_METHOD

METHOD CALL_STACK_LOADPOS
VAR_IN_OUT
	LRCYCPOS : LREAL;
	LRLOADPOS : LREAL;
END_VAR
END_METHOD

METHOD CALL_STACK_TAKEPOS
VAR_IN_OUT
	LRCYCPOS : LREAL;
END_VAR
END_METHOD

METHOD FUN_PERIODCNTRDIFF : LREAL
VAR_INPUT
	UIDIFF : UINT;
END_VAR
VAR_OUTPUT
	IOUT : INT;
END_VAR
END_METHOD

METHOD GET_LRLATESTDIST : LREAL
VAR_IN_OUT
	LRCYCPOS : LREAL;
END_VAR
END_METHOD

METHOD GET_LRTAKEPOS : LREAL
VAR_IN_OUT
	LRCYCPOS : LREAL;
END_VAR
END_METHOD

METHOD REVOKETAKEPOS
END_METHOD

METHOD SET_CYCSETPOS
VAR_IN_OUT
	LRCYCPOS : LREAL;
END_VAR
END_METHOD

METHOD SET_TPPOS
VAR_IN_OUT
	LRCYCPOS : LREAL;
	LRLOADTPPOS : LREAL;
END_VAR
END_METHOD

(* ---- L_MB1P_TPAVERAGEDIFF.fb ---- *)
FUNCTION_BLOCK L_MB1P_TPAVERAGEDIFF
VAR_INPUT
	XENABLE : BOOL;
	BYNROFCYCLES : BYTE := 20;
	XTPRECEIVED : BOOL;
	LRSETTPDIFFERENCE : LREAL;
	XTPERRORLIMITED : BOOL;
	LRSETMARKDISTANCE : LREAL;
	LRSETMAXAVERAGE : LREAL := 100;
END_VAR
VAR_OUTPUT
	LRTPERRORAVERAGE : LREAL;
	XAVERAGELIMITED : BOOL;
	LROPTIMISEDGEARFACTOR : LREAL;
END_VAR
VAR
	LRPROCENT : LREAL;
	BYNROFCYCLESINTERNAL : BYTE;
	XTPRECEIVEDOLD : BOOL;
	LRTOTALERROR : LREAL;
	BYCOUNTER : BYTE;
	LROPTIMIZATIONUNCLAMPED : LREAL;
END_VAR
END_FUNCTION_BLOCK
